// ---- 99_Test/PRG_TestPeakLive.TcPOU
PROGRAM PRG_TestPeakLive		// 피크컷(3)·통합(4) 모드 실제 경로 시험 (시험 모드, MAIN이 부름). bStart := TRUE로 시작, 약 10~15분
// 부하 모델: 가상 접속점 P = ESS 출력 − 부하 (수전 = 부하 − ESS 방전). 목표 피크 300 kW, 방전 허용 시간 끔 (PLC 시계 UTC)
// 피크컷: P1 부하 500 → 피크 방전, P2 부하 200 → 0, P3 자동 충전 시간 → 충전, P4 잔량 방전 시간 → 방전 (역송 방지 상한)
// 통합:   I1 부하 200·시간표 +100 → 100, I2 부하 600 → 피크·시간표 중 큰 값, I3 부하 200·시간표 −200 → 충전, I4 잔량 방전
// 구간마다 조건이 5 s 이어지면 통과·기록. 끝나면 설정·가상신호·운전 모드 되돌리고 PCS 정지
VAR
	bStart		: BOOL;				// TRUE로 쓰면 시작
	bDone		: BOOL;
	bPass		: BOOL;				// 8구간 모두 통과
	nStep		: UINT;
	wsStep		: WSTRING(80);		// 지금 단계
	wsFail		: WSTRING(80);
	(* 지금 값 *)
	fLoadSim	: REAL;				// kW, 모의 부하
	fImport		: REAL;				// kW, 수전 (= 부하 − ESS 출력)
	nActiveMode	: UINT;				// 3 = 피크컷, 4 = 통합
	nState		: UINT;				// 켜진 모드 상태 (GVL_CM_RSN: 0 정상, 11 피크, 12 피크 필요 없음, 13 자동 충전, 14 잔량 방전, 15 스케줄·피크, 6 역송 방지)
	fModeP		: REAL;				// 모드가 낸 값 (kW, 방전 +)
	fMgrP		: REAL;				// 관리자 지령
	fUnitP		: REAL;				// 가상 PCS 실제 출력
	fPeakCtrl	: REAL;				// 피크 제어량
	nRemainMin	: UINT;				// 15분 구간 남은 분
	fSoc		: REAL;				// %
	eRun		: E_RunState;
	stNow		: ST_LocalTime;
	(* 구간 결과 (통과 때 실제 출력 kW) *)
	bP1Peak		: BOOL;		fP1		: REAL;		// 피크컷: 부하 500 → 피크 방전
	bP2Below	: BOOL;		fP2		: REAL;		// 피크컷: 부하 200 → 0
	bP3AutoChg	: BOOL;		fP3		: REAL;		// 피크컷: 자동 충전
	bP4Remain	: BOOL;		fP4		: REAL;		// 피크컷: 잔량 방전
	bI1Sched	: BOOL;		fI1		: REAL;		// 통합: 시간표 +100
	bI2Peak		: BOOL;		fI2		: REAL;		// 통합: 피크·시간표 중 큰 값
	bI3Chg		: BOOL;		fI3		: REAL;		// 통합: 시간표 충전 −200
	bI4Remain	: BOOL;		fI4		: REAL;		// 통합: 잔량 방전
	(* 내부 *)
	bLoadSim	: BOOL;
	nLastStep	: UINT;
	tonStep		: TON;
	tonOk		: TON;
	bCond		: BOOL;
	bBackedUp	: BOOL;
	stCommonBak	: ST_CmCommonSet;
	stSchedBak	: ST_CmScheduleSet;
	stPeakBak	: ST_CmPeakCutSet;
	stSPBak		: ST_CmSchedPeakSet;
	stVirtBak	: ST_VirtualSet;
	stCmBak		: ST_CtrlModeSet;
	stMgrOut	: ST_SourceOutput;
	nMin		: UINT;
	nSeason		: UINT;
	k			: UINT;
	nWinStart	: UINT;		// HHMM
	nWinEnd		: UINT;		// HHMM (지금 + 3분)
	nSlotEnd	: UINT;		// HHMM (지금 + 30분)
END_VAR

// 지금 값
stNow		:= MAIN.fbClock.q_stTime;
nActiveMode	:= GVL_SITE.g_fbCtrlMode1.q_nActive;
stMgrOut	:= GVL_SITE.g_fbCtrlMode1.Output;
fMgrP		:= stMgrOut.fPSet;	// [16번 수정 2026-11-09: 관리자가 접속점 그룹 단위 → 접속점 그룹 지령 칸. 원래 stMgrOut.astUnit[1].fPSet (PCS2는 Manual이라 접속점 그룹 지령이 유닛 1로 감)]
fUnitP		:= MAIN.fbSnapshot.q_astUnit[1].stP.fValue;
eRun		:= MAIN.fbSnapshot.q_astUnit[1].eRunState;
fSoc		:= MAIN.fbGroupView.q_astView[1].stSocAvg.fValue;
IF nActiveMode = 4 THEN
	nState		:= GVL_SITE.g_fbCmSchedPeak1.q_nState;
	fModeP		:= GVL_SITE.g_fbCmSchedPeak1.q_fOutP;
	fPeakCtrl	:= GVL_SITE.g_fbCmSchedPeak1.q_fPeakCtrl;
	nRemainMin	:= GVL_SITE.g_fbCmSchedPeak1.q_nRemainMin;
ELSE
	nState		:= GVL_SITE.g_fbCmPeakCut1.q_nState;
	fModeP		:= GVL_SITE.g_fbCmPeakCut1.q_fOutP;
	fPeakCtrl	:= GVL_SITE.g_fbCmPeakCut1.q_fPeakCtrl;
	nRemainMin	:= GVL_SITE.g_fbCmPeakCut1.q_nRemainMin;
END_IF
// 부하 모델: 접속점 P (공급 +) = ESS 출력 − 부하
IF bLoadSim THEN
	GVL_TEST.g_astVirtual[1].bPEna	:= TRUE;
	GVL_TEST.g_astVirtual[1].fP		:= MAIN.fbGroupView.q_astView[1].fPOut - fLoadSim;	// 그룹 출력 (PCS2는 Manual 0)
END_IF
fImport := fLoadSim - fUnitP;
// 시간 구간 (지금 분 ~ +3분, 시간표 칸은 +30분)
nMin		:= stNow.nHour * 60 + stNow.nMinute;
nWinStart	:= (nMin / 60) * 100 + nMin MOD 60;
nWinEnd		:= (((nMin + 3) MOD 1440) / 60) * 100 + ((nMin + 3) MOD 1440) MOD 60;
nSlotEnd	:= (((nMin + 30) MOD 1440) / 60) * 100 + ((nMin + 30) MOD 1440) MOD 60;

tonStep(IN := nStep >= 20 AND nStep < 900, PT := T#240S);
bCond := FALSE;

CASE nStep OF
	0:
		IF bStart THEN
			bStart := FALSE;	bDone := FALSE;	bPass := FALSE;	wsFail := "";
			bP1Peak := FALSE;	bP2Below := FALSE;	bP3AutoChg := FALSE;	bP4Remain := FALSE;
			bI1Sched := FALSE;	bI2Peak := FALSE;	bI3Chg := FALSE;	bI4Remain := FALSE;
			nStep := 10;
		ELSIF NOT bDone THEN
			wsStep := "대기: bStart := TRUE로 시작";
		END_IF

	10:	// 준비
		wsStep := "설정 준비";
		IF NOT stNow.bValid OR stNow.nMonth < 1 OR stNow.nMonth > 12 OR stNow.nDay < 1 OR stNow.nDay > 31 OR stNow.nDayOfWeek > 6 THEN
			wsFail := "PLC 시각 무효";
			nStep := 900;
		ELSIF nMin + 40 >= 1440 THEN
			wsFail := "자정 가까움: 40분 뒤 다시";
			nStep := 900;
		ELSE
			stCommonBak	:= GVL_PERSIST.g_stModuleSet.stCmCommon;
			stSchedBak	:= GVL_PERSIST.g_stModuleSet.stCmSchedule1;
			stPeakBak	:= GVL_PERSIST.g_stModuleSet.stCmPeakCut1;
			stSPBak		:= GVL_PERSIST.g_stModuleSet.stCmSchedPeak1;
			stVirtBak	:= GVL_TEST.g_astVirtual[1];
			stCmBak		:= GVL_PERSIST.g_stModuleSet.stCtrlMode1;
			GVL_PERSIST.g_stModuleSet.stCtrlMode1.ePccShare := E_PccShare.Actual;	// PCS1이 접속점 실측 그대로 (PCS2는 Manual 0)
			bBackedUp	:= TRUE;
			GVL_PERSIST.g_stModuleSet.stCmCommon.stDis.bUse := FALSE;
			GVL_PERSIST.g_stModuleSet.stCmCommon.abHoliday[stNow.nMonth, stNow.nDay] := FALSE;
			GVL_PERSIST.g_stModuleSet.stCmPeakCut1.stPeak.fTarget	:= 300.0;
			GVL_PERSIST.g_stModuleSet.stCmPeakCut1.stAutoChg.bUse	:= FALSE;
			GVL_PERSIST.g_stModuleSet.stCmPeakCut1.stRemain.bUse		:= FALSE;
			GVL_PERSIST.g_stModuleSet.stCmSchedPeak1.stPeak.fTarget	:= 300.0;
			GVL_PERSIST.g_stModuleSet.stCmSchedPeak1.stRemain.bUse	:= FALSE;
			nSeason := GVL_PERSIST.g_stModuleSet.stCmCommon.anSeasonOfMonth[stNow.nMonth];
			IF nSeason > 2 THEN
				nSeason := 0;
			END_IF
			FOR k := 1 TO GVL_PARAM.SCHED_SLOT_COUNT DO
				GVL_PERSIST.g_stModuleSet.stCmSchedule1.astSlot[nSeason, stNow.nDayOfWeek, k].nStart	:= 0;
				GVL_PERSIST.g_stModuleSet.stCmSchedule1.astSlot[nSeason, stNow.nDayOfWeek, k].nEnd	:= 0;
				GVL_PERSIST.g_stModuleSet.stCmSchedule1.astSlot[nSeason, stNow.nDayOfWeek, k].fP		:= 0.0;
			END_FOR
			fLoadSim	:= 500.0;
			bLoadSim	:= TRUE;
			GVL_PERSIST.g_aeOpMode[1] := E_OpMode.Auto;
			nStep := 20;
		END_IF

	20:
		wsStep := "Auto 전환 대기";
		IF MAIN.fbModeSwitch.q_aeOpMode[1] = E_OpMode.Auto THEN
			GVL_SITE.g_fbSrcTest.i_nBatGroup	:= 0;
			GVL_SITE.g_fbSrcTest.i_eBatReq		:= E_BatCmd.Close;
			nStep := 30;
		END_IF
	30:
		wsStep := "배터리 투입 대기";
		IF MAIN.fbBatGroup.q_astBatGroup[1].bReady THEN
			GVL_SITE.g_fbSrcTest.i_nPcsUnit	:= 0;
			GVL_SITE.g_fbSrcTest.i_ePcsReq	:= E_PcsCmd.Run;
			nStep := 40;
		END_IF
	40:
		wsStep := "PCS Run 대기";
		IF eRun = E_RunState.Run THEN
			GVL_SITE.g_fbCtrlMode1.i_nModeReq := 3;
			nStep := 50;
		END_IF
	50:
		wsStep := "피크컷 모드 켜는 중";
		IF nActiveMode = 3 THEN
			nStep := 100;
		END_IF

	100: // P1 부하 500 > 목표 300 → 피크 방전
		wsStep := "P1 피크컷: 부하 500 > 목표 300";
		bCond := nActiveMode = 3 AND nState = GVL_CM_RSN.PEAK AND fPeakCtrl > 0.0 AND fModeP > 0.0 AND ABS(fUnitP - fModeP) < 5.0;
		IF tonOk.Q THEN
			bP1Peak := TRUE;	fP1 := fUnitP;
			fLoadSim := 200.0;
			nStep := 110;
		END_IF
	110: // P2 부하 200 < 목표 → 0
		wsStep := "P2 피크컷: 부하 200 < 목표 300";
		bCond := nState = GVL_CM_RSN.BELOW_PEAK AND ABS(fUnitP) < 5.0;
		IF tonOk.Q THEN
			bP2Below := TRUE;	fP2 := fUnitP;
			GVL_PERSIST.g_stModuleSet.stCmPeakCut1.stAutoChg.nStart	:= nWinStart;
			GVL_PERSIST.g_stModuleSet.stCmPeakCut1.stAutoChg.nEnd	:= nWinEnd;
			GVL_PERSIST.g_stModuleSet.stCmPeakCut1.stAutoChg.fSoc	:= 100.0;
			GVL_PERSIST.g_stModuleSet.stCmPeakCut1.stAutoChg.bUse	:= TRUE;
			nStep := 120;
		END_IF
	120: // P3 자동 충전 시간
		wsStep := "P3 피크컷: 자동 충전 시간";
		bCond := nState = GVL_CM_RSN.AUTO_CHG AND fModeP < -5.0 AND fUnitP < -5.0;
		IF tonOk.Q THEN
			bP3AutoChg := TRUE;	fP3 := fUnitP;
			GVL_PERSIST.g_stModuleSet.stCmPeakCut1.stAutoChg.bUse	:= FALSE;
			GVL_PERSIST.g_stModuleSet.stCmPeakCut1.stRemain.nStart	:= nWinStart;
			GVL_PERSIST.g_stModuleSet.stCmPeakCut1.stRemain.nEnd		:= nWinEnd;
			GVL_PERSIST.g_stModuleSet.stCmPeakCut1.stRemain.fSoc		:= 10.0;
			GVL_PERSIST.g_stModuleSet.stCmPeakCut1.stRemain.bUse		:= TRUE;
			fLoadSim := 500.0;
			nStep := 130;
		END_IF
	130: // P4 잔량 방전 시간 (역송 방지 상한)
		wsStep := "P4 피크컷: 잔량 방전 시간";
		bCond := (nState = GVL_CM_RSN.REMAIN_DIS OR nState = GVL_CM_RSN.REV_LIMIT) AND fModeP > 5.0 AND ABS(fUnitP - fModeP) < 5.0 AND fUnitP < fLoadSim;
		IF tonOk.Q THEN
			bP4Remain := TRUE;	fP4 := fUnitP;
			GVL_PERSIST.g_stModuleSet.stCmPeakCut1.stRemain.bUse := FALSE;
			// 통합 준비: 시간표 +100 (지금 ~ +30분), 부하 200
			GVL_PERSIST.g_stModuleSet.stCmSchedule1.astSlot[nSeason, stNow.nDayOfWeek, 1].nStart	:= nWinStart;
			GVL_PERSIST.g_stModuleSet.stCmSchedule1.astSlot[nSeason, stNow.nDayOfWeek, 1].nEnd	:= nSlotEnd;
			GVL_PERSIST.g_stModuleSet.stCmSchedule1.astSlot[nSeason, stNow.nDayOfWeek, 1].fP		:= 100.0;
			fLoadSim := 200.0;
			GVL_SITE.g_fbCtrlMode1.i_nModeReq := 4;
			nStep := 200;
		END_IF

	200:
		wsStep := "통합 모드 켜는 중";
		IF nActiveMode = 4 THEN
			nStep := 210;
		END_IF
	210: // I1 부하 200 (피크 아님) → 시간표 +100
		wsStep := "I1 통합: 부하 200, 시간표 +100";
		bCond := nState = 0 AND ABS(fModeP - 100.0) < 0.5 AND ABS(fUnitP - 100.0) < 5.0;
		IF tonOk.Q THEN
			bI1Sched := TRUE;	fI1 := fUnitP;
			fLoadSim := 600.0;
			nStep := 220;
		END_IF
	220: // I2 부하 600 > 목표 → 피크 제어량과 시간표 중 큰 값
		wsStep := "I2 통합: 부하 600 > 목표 300";
		bCond := nState = GVL_CM_RSN.SCHED_PEAK AND fPeakCtrl > 0.0 AND fModeP >= 99.9 AND ABS(fModeP - MAX(fPeakCtrl, 100.0)) < 0.5 AND ABS(fUnitP - fModeP) < 5.0;
		IF tonOk.Q THEN
			bI2Peak := TRUE;	fI2 := fUnitP;
			GVL_PERSIST.g_stModuleSet.stCmSchedule1.astSlot[nSeason, stNow.nDayOfWeek, 1].fP := -200.0;
			fLoadSim := 200.0;
			nStep := 230;
		END_IF
	230: // I3 부하 200, 시간표 충전 −200
		wsStep := "I3 통합: 부하 200, 시간표 -200";
		bCond := nState = 0 AND ABS(fModeP + 200.0) < 0.5 AND ABS(fUnitP + 200.0) < 5.0;
		IF tonOk.Q THEN
			bI3Chg := TRUE;	fI3 := fUnitP;
			GVL_PERSIST.g_stModuleSet.stCmSchedPeak1.stRemain.nStart	:= nWinStart;
			GVL_PERSIST.g_stModuleSet.stCmSchedPeak1.stRemain.nEnd	:= nWinEnd;
			GVL_PERSIST.g_stModuleSet.stCmSchedPeak1.stRemain.fSoc	:= 10.0;
			GVL_PERSIST.g_stModuleSet.stCmSchedPeak1.stRemain.bUse	:= TRUE;
			fLoadSim := 500.0;
			nStep := 240;
		END_IF
	240: // I4 잔량 방전
		wsStep := "I4 통합: 잔량 방전 시간";
		bCond := (nState = GVL_CM_RSN.REMAIN_DIS OR nState = GVL_CM_RSN.REV_LIMIT) AND fModeP > 5.0 AND ABS(fUnitP - fModeP) < 5.0 AND fUnitP < fLoadSim;
		IF tonOk.Q THEN
			bI4Remain := TRUE;	fI4 := fUnitP;
			nStep := 900;
		END_IF

	900: // 정리
		GVL_SITE.g_fbCtrlMode1.i_nModeReq	:= 0;
		GVL_SITE.g_fbSrcTest.i_nPcsUnit		:= 0;
		GVL_SITE.g_fbSrcTest.i_ePcsReq		:= E_PcsCmd.Stop;
		bLoadSim := FALSE;
		IF bBackedUp THEN
			GVL_PERSIST.g_stModuleSet.stCmCommon	:= stCommonBak;
			GVL_PERSIST.g_stModuleSet.stCmSchedule1	:= stSchedBak;
			GVL_PERSIST.g_stModuleSet.stCmPeakCut1	:= stPeakBak;
			GVL_PERSIST.g_stModuleSet.stCmSchedPeak1	:= stSPBak;
			GVL_TEST.g_astVirtual[1]				:= stVirtBak;
			GVL_PERSIST.g_stModuleSet.stCtrlMode1	:= stCmBak;
			bBackedUp := FALSE;
		END_IF
		GVL_PERSIST.g_aeOpMode[1] := E_OpMode.Manual;
		bPass := bP1Peak AND bP2Below AND bP3AutoChg AND bP4Remain AND bI1Sched AND bI2Peak AND bI3Chg AND bI4Remain AND wsFail = "";
		bDone := TRUE;
		IF bPass THEN
			wsStep := "끝: 통과";
		ELSE
			wsStep := "끝: 실패 (wsFail·구간 결과 확인)";
		END_IF
		nStep := 0;
END_CASE

// 조건이 5 s 이어지면 통과 (단계가 바뀌면 다시 셈)
tonOk(IN := bCond AND nStep = nLastStep, PT := T#5S);
IF tonStep.Q AND nStep >= 20 AND nStep < 900 THEN
	wsFail	:= WCONCAT("시간 초과: ", wsStep);
	nStep	:= 900;
END_IF
IF nStep <> nLastStep THEN
	tonStep(IN := FALSE);
	tonOk(IN := FALSE);
	nLastStep := nStep;
END_IF

END_PROGRAM

// ---- 99_Test/PRG_TestUnitMode.TcPOU
PROGRAM PRG_TestUnitMode		// PCS별(유닛 단위) 제어 모드 자동 시험 (GVL_SITE.TEST_MODE일 때 MAIN이 부름). 따로 둔 인스턴스만 씀 (장비 지령에 영향 없음)
// 온라인에서 bDone = TRUE가 되면 fbTally.q_nPass·q_nFail, 실패하면 fbTally.q_anFail. bRestart := TRUE로 다시 돌림
// 40~41: 유닛 단위 출력 칸, 42~44: 접속점 몫 (ByRating·Actual·Fixed), 45~47: 설정 점검, 48~50: FB_UnitView 버스 몫, 51~57: 스탠다드 스케줄 모드, 58~63: NaN·무한대 거르기 (PLC가 멈추지 않아야 함)
VAR
	bRestart	: BOOL;
	bDone		: BOOL;
	nStep		: UINT;
	fbTally		: FB_TestTally;
	fbConstU	: FB_CmConstPower	:= (i_nModuleId := 9012, i_sName := 'TestConstU');
	fbMgrU		: FB_CtrlModeMgr	:= (i_nModuleId := 9010, i_sName := 'TestMgrU', i_nUnit := 1);
	aipMode		: ARRAY[1..GVL_PARAM.CTRL_MODE_COUNT] OF I_ControlMode;
	astUv		: ARRAY[1..GVL_PARAM.UNIT_COUNT] OF ST_UnitView;	// 관리자에 주소로 넘기는 유닛 값 (시험이 채움)
	stGrpView	: ST_GroupView;			// 지령원 공통 입력 (유닛 단위에서는 안 봄)
	stReg		: ST_SourceReg := (bEnable := TRUE, nGrade := 1, ePowerMode := E_SourceMode.Auto, nGroup := 0, tExpire := T#10S);
	stMgrOut	: ST_SourceOutput;
	wsTmp		: WSTRING(63);
	(* FB_UnitView 시험 (유닛 1 기준, 유닛이 2개 이상이면 유닛 2도) *)
	fbUv		: FB_UnitView;
	astView		: ARRAY[1..GVL_PARAM.GROUP_COUNT] OF ST_GroupView;
	astUnit		: ARRAY[1..GVL_PARAM.UNIT_COUNT] OF ST_UnitState;
	astAvail	: ARRAY[1..GVL_PARAM.UNIT_COUNT] OF ST_UnitAvail;
	astCfg		: ARRAY[1..GVL_PARAM.UNIT_COUNT] OF ST_UnitCfg;
	astEnv		: ARRAY[1..GVL_PARAM.UNIT_COUNT] OF ST_UnitEnvelope;
	astBat		: ARRAY[1..GVL_PARAM.BAT_COUNT] OF ST_BatGroupState;
	astBatEnv	: ARRAY[1..GVL_PARAM.BAT_COUNT] OF ST_BatEnvelope;
	fShareExp	: REAL;
	(* 스탠다드 스케줄 모드 시험 *)
	fbStd		: FB_CmStdSchedule	:= (i_nModuleId := 9013, i_sName := 'TestStdSched');
	stStdView	: ST_CtrlModeView;
	stStdOut	: ST_CtrlModeOut;
	nInfBits	: DWORD := 16#7F800000;	// +무한대 비트 (NaN은 크기 비교에서 부동소수점 예외로 PLC가 멈추므로 시험에 쓰지 않음)
	fInf		: REAL;
	nBad0		: UDINT;
	nNanBits	: DWORD := 16#7FC00000;	// NaN 비트 (거르기 시험: 비교하기 전에 걸러져야 PLC가 멈추지 않음)
	fNan		: REAL;
	fbEmsCmd	: FB_EmsCommand;		// EMS 명령 핸들러 시험 인스턴스
	astPcsRx	: ARRAY[0..GVL_PARAM.PCS_COUNT - 1] OF ST_MqttCommand_Rx;
	astBatRx	: ARRAY[0..GVL_PARAM.BMS_COUNT - 1] OF ST_MqttCommand_Rx;
	nPSeq0		: UDINT;
	nRunSeq0	: UDINT;		// 시험 전 이상값 버린 수 (누계라 다시 돌려도 맞게)
	u			: UINT;
END_VAR

IF bRestart THEN
	bRestart	:= FALSE;
	bDone		:= FALSE;
	nStep		:= 0;
END_IF

CASE nStep OF
	0:	// 준비: 정출력 80 kW 하나, 유닛 1 값 (출력 100, 그룹 출력 300, 접속점 -200 = 수전 200 → 그룹 부하 500, 몫 0.5)
		fbTally.M_Reset();
		aipMode[1]					:= fbConstU;
		fbConstU.i_stSet.fPSet		:= 80.0;
		fbConstU.i_stSet.bQSet		:= FALSE;
		fbConstU.i_stSet.tDuration	:= T#0S;
		astUv[1].nUnit				:= 1;
		astUv[1].bAvail				:= TRUE;
		astUv[1].stView.nUnitAvail	:= 1;
		astUv[1].stView.fPRatedAvail	:= 1000.0;
		astUv[1].stView.fPOut		:= 100.0;
		astUv[1].stView.stPcc.stMeas.stP.bValid	:= TRUE;
		astUv[1].stView.stPcc.stMeas.stP.fValue	:= -200.0;
		astUv[1].fGroupPOut			:= 300.0;
		astUv[1].fRatingShare		:= 0.5;
		fbMgrU.i_aipMode			:= aipMode;
		fbMgrU.i_stSet.bZeroOnSwitch	:= TRUE;
		fbMgrU.i_stSet.tZeroDelay	:= T#1S;
		fbMgrU.i_stSet.nFallback	:= 0;
		fbMgrU.i_stSet.ePccShare	:= E_PccShare.ByRating;
		fbMgrU.i_stSet.fPccRatio	:= 1.0;
		fbMgrU.i_pUnitView			:= ADR(astUv);
		wsTmp := fbMgrU.M_CheckSet();
		fbTally.M_Check(i_nId := 40, i_bOk := wsTmp = "");
		fbMgrU.i_nModeReq := 1;
		nStep := 10;

	10:	// 정출력 진입: 유닛 1 칸에만 80, 그룹 지령은 없음. 몫 0.5 → 모드가 본 접속점 = 100 - 0.5 × 500 = -150
		A_Cycle();
		fbTally.M_Check(i_nId := 41, i_bOk := fbMgrU.q_nActive = 1 AND stMgrOut.astUnit[1].bPSetActive AND ABS(stMgrOut.astUnit[1].fPSet - 80.0) < 0.01 AND NOT stMgrOut.bPSetActive);
		fbTally.M_Check(i_nId := 42, i_bOk := ABS(fbMgrU.q_fPccP + 150.0) < 0.01);
		fbMgrU.i_stSet.ePccShare := E_PccShare.Actual;
		nStep := 11;

	11:	// Actual: 실측 그대로 -200
		A_Cycle();
		fbTally.M_Check(i_nId := 43, i_bOk := ABS(fbMgrU.q_fPccP + 200.0) < 0.01);
		fbMgrU.i_stSet.ePccShare := E_PccShare.Fixed;
		fbMgrU.i_stSet.fPccRatio := 0.2;
		nStep := 12;

	12:	// Fixed 0.2: 100 - 0.2 × 500 = 0
		A_Cycle();
		fbTally.M_Check(i_nId := 44, i_bOk := ABS(fbMgrU.q_fPccP) < 0.01);
		// 설정 점검: 몫 범위 밖, 유닛 값 연결 안 됨, 유닛 번호 범위 밖
		fbMgrU.i_stSet.fPccRatio := 1.5;
		wsTmp := fbMgrU.M_CheckSet();
		fbTally.M_Check(i_nId := 45, i_bOk := wsTmp <> "");
		fbMgrU.i_stSet.fPccRatio := 0.2;
		fbMgrU.i_pUnitView := 0;
		wsTmp := fbMgrU.M_CheckSet();
		fbTally.M_Check(i_nId := 46, i_bOk := wsTmp <> "");
		fbMgrU.i_pUnitView := ADR(astUv);
		fbMgrU.i_nUnit := GVL_PARAM.UNIT_COUNT + 1;
		wsTmp := fbMgrU.M_CheckSet();
		fbTally.M_Check(i_nId := 47, i_bOk := wsTmp <> "");
		fbMgrU.i_nUnit := 1;
		A_UnitViewTest();
		A_StdScheduleTest();
		A_NanTest();
		nStep := 99;

	99:
		bDone := TRUE;
END_CASE

ACTION A_Cycle:
fbMgrU.i_pUnitView := ADR(astUv);	// 온라인 변경 뒤에도 맞게 매번
fbMgrU.M_Cycle(i_stReg := stReg, i_stView := stGrpView);
stMgrOut := fbMgrU.Output;
END_ACTION

ACTION A_UnitViewTest:
// FB_UnitView: 그룹 1 (접속점 -200, 그룹 출력 300, 가용 한도 합 2000), 버스 1 (방전 한도 1200, 충전 한도 800, 용량 4000, SOC 60)
// 유닛 1 정격 1000 (한도 1000, 출력 100). 유닛이 2개 이상이면 유닛 2도 같은 버스·정격 1000 → 버스 몫 0.5, 아니면 1
astView[1].stPcc.stMeas.stP.bValid	:= TRUE;
astView[1].stPcc.stMeas.stP.fValue	:= -200.0;
astView[1].fPOut			:= 300.0;
astView[1].fPRatedAvail		:= 2000.0;
astBat[1].bUsable			:= TRUE;
astBat[1].fCapacity			:= 4000.0;
astBat[1].stSoc.bValid		:= TRUE;
astBat[1].stSoc.fValue		:= 60.0;
astBatEnv[1].stP.fMax		:= 1200.0;
astBatEnv[1].stP.fMin		:= -800.0;
FOR u := 1 TO GVL_PARAM.UNIT_COUNT DO
	astCfg[u].nGroup		:= 1;
	astCfg[u].nBatGroup		:= 1;
	astCfg[u].fPRated		:= 1000.0;
	astCfg[u].fQRated		:= 500.0;
	astAvail[u].bAvail		:= TRUE;
	astEnv[u].stP.fMax		:= 1000.0;
	astEnv[u].stQ.fMax		:= 500.0;
	astUnit[u].stP.bValid	:= TRUE;
	astUnit[u].stP.fValue	:= 100.0;
END_FOR
fShareExp := 1.0 / UINT_TO_REAL(GVL_PARAM.UNIT_COUNT);
fbUv(iq_astView := astView, iq_astUnit := astUnit, iq_astAvail := astAvail, iq_astUnitCfg := astCfg,
	iq_astUnitEnv := astEnv, iq_astBatGroup := astBat, iq_astBatEnv := astBatEnv);
// 48) 유닛 1: 출력·한도·접속점·그룹 출력·정격 몫 (1000 / 2000)
fbTally.M_Check(i_nId := 48, i_bOk := fbUv.q_astView[1].stView.nUnitAvail = 1 AND ABS(fbUv.q_astView[1].stView.fPOut - 100.0) < 0.01
	AND ABS(fbUv.q_astView[1].stView.fPRatedAvail - 1000.0) < 0.01 AND ABS(fbUv.q_astView[1].stView.stPcc.stMeas.stP.fValue + 200.0) < 0.01
	AND ABS(fbUv.q_astView[1].fGroupPOut - 300.0) < 0.01 AND ABS(fbUv.q_astView[1].fRatingShare - 0.5) < 0.001);
// 49) 버스 몫: 용량·방전·충전 한도 × 몫, SOC 그대로
fbTally.M_Check(i_nId := 49, i_bOk := ABS(fbUv.q_astView[1].stView.fCapacity - 4000.0 * fShareExp) < 0.1
	AND ABS(fbUv.q_astView[1].stView.fPDisMax - MIN(1200.0 * fShareExp, 1000.0)) < 0.1 AND ABS(fbUv.q_astView[1].stView.fPChgMax - MIN(800.0 * fShareExp, 1000.0)) < 0.1
	AND fbUv.q_astView[1].stView.stSocAvg.bValid AND ABS(fbUv.q_astView[1].stView.stSocAvg.fValue - 60.0) < 0.01);
// 50) 가용이 아닌 유닛: 가용 0, 몫 0, 용량 0
astAvail[1].bAvail := FALSE;
fbUv(iq_astView := astView, iq_astUnit := astUnit, iq_astAvail := astAvail, iq_astUnitCfg := astCfg,
	iq_astUnitEnv := astEnv, iq_astBatGroup := astBat, iq_astBatEnv := astBatEnv);
fbTally.M_Check(i_nId := 50, i_bOk := fbUv.q_astView[1].stView.nUnitAvail = 0 AND fbUv.q_astView[1].fRatingShare = 0.0 AND fbUv.q_astView[1].stView.fCapacity = 0.0
	AND ABS(fbUv.q_astView[1].stView.fPOut - 100.0) < 0.01);
astAvail[1].bAvail := TRUE;
END_ACTION

ACTION A_StdScheduleTest:
// 스탠다드 스케줄: EMS가 9시 방전 100, 10시 정지를 보내는 흐름 (한 스캔씩 직접 부름)
stStdView.stGroup.nUnitAvail := 1;
// 켜지기 전에 온 지령(번호 5, 50 kW)은 쓰지 않음
fbStd.i_astCmd[1].bUse		:= TRUE;	// [16번 수정 2026-11-09: 모드가 유닛마다 칸을 받음 (유닛 1 칸으로 시험). 원래 fbStd.i_stCmd, 출력 stStdOut.bPSetActive·fPSet]
fbStd.i_astCmd[1].bAlive	:= TRUE;
fbStd.i_astCmd[1].nPSeq		:= 5;
fbStd.i_astCmd[1].fP		:= 50.0;
fbStd.i_astCmd[1].nStateSeq	:= 3;
fbStd.i_astCmd[1].eState	:= E_PcsCmd.Run;
fbStd.M_Enter(i_stView := stStdView);
stStdOut := fbStd.M_Calc(i_stView := stStdView);
fbTally.M_Check(i_nId := 51, i_bOk := stStdOut.bUnitOut AND stStdOut.astUnit[1].bPSetActive AND stStdOut.astUnit[1].fPSet = 0.0 AND fbStd.q_nState = 3 AND NOT fbStd.q_abHold[1]);
// 9시: 방전 100 → 100, 다음 지령까지 유지
fbStd.i_astCmd[1].nPSeq	:= 6;
fbStd.i_astCmd[1].fP	:= 100.0;
stStdOut := fbStd.M_Calc(i_stView := stStdView);
stStdOut := fbStd.M_Calc(i_stView := stStdView);
fbTally.M_Check(i_nId := 52, i_bOk := ABS(stStdOut.astUnit[1].fPSet - 100.0) < 0.01 AND fbStd.q_nState = 0 AND fbStd.q_nCmdCount = 1);
// 10시: 정지 → 0 (새 P 지령 대기)
fbStd.i_astCmd[1].nStateSeq	:= 4;
fbStd.i_astCmd[1].eState	:= E_PcsCmd.Stop;
stStdOut := fbStd.M_Calc(i_stView := stStdView);
fbTally.M_Check(i_nId := 53, i_bOk := stStdOut.astUnit[1].bPSetActive AND stStdOut.astUnit[1].fPSet = 0.0 AND fbStd.q_nState = 3);
// Run만 다시 와도 옛 100은 되살아나지 않음
fbStd.i_astCmd[1].nStateSeq	:= 5;
fbStd.i_astCmd[1].eState	:= E_PcsCmd.Run;
stStdOut := fbStd.M_Calc(i_stView := stStdView);
fbTally.M_Check(i_nId := 54, i_bOk := stStdOut.astUnit[1].fPSet = 0.0 AND NOT fbStd.q_abHold[1]);
// 충전 -200 → -200. 이상값(무한대)은 버리고 앞 값 유지
fbStd.i_astCmd[1].nPSeq	:= 7;
fbStd.i_astCmd[1].fP	:= -200.0;
stStdOut := fbStd.M_Calc(i_stView := stStdView);
nBad0 := fbStd.q_nBadCount;
fbStd.i_astCmd[1].nPSeq	:= 8;
MEMCPY(destAddr := ADR(fInf), srcAddr := ADR(nInfBits), n := SIZEOF(fInf));	// +무한대 (비트로 만듦)
fbStd.i_astCmd[1].fP	:= fInf;
stStdOut := fbStd.M_Calc(i_stView := stStdView);
fbTally.M_Check(i_nId := 55, i_bOk := ABS(stStdOut.astUnit[1].fPSet + 200.0) < 0.01 AND fbStd.q_nBadCount = nBad0 + 1);
// EMS 끊김 → 0, 돌아와도 옛 값은 되살아나지 않음
fbStd.i_astCmd[1].bAlive := FALSE;
stStdOut := fbStd.M_Calc(i_stView := stStdView);
fbTally.M_Check(i_nId := 56, i_bOk := stStdOut.astUnit[1].fPSet = 0.0 AND fbStd.q_nState = 2);
fbStd.i_astCmd[1].bAlive := TRUE;
stStdOut := fbStd.M_Calc(i_stView := stStdView);
fbTally.M_Check(i_nId := 57, i_bOk := stStdOut.astUnit[1].fPSet = 0.0 AND fbStd.q_nState = 3);
fbStd.M_Exit();
END_ACTION

ACTION A_NanTest:
// NaN·무한대: 비트로 먼저 거르는지 (거르지 못하면 여기서 PLC가 멈춤)
MEMCPY(destAddr := ADR(fNan), srcAddr := ADR(nNanBits), n := SIZEOF(fNan));
// 58) F_IsFinite: NaN·무한대 FALSE, 보통 숫자 TRUE
fbTally.M_Check(i_nId := 58, i_bOk := NOT F_IsFinite(fNan) AND NOT F_IsFinite(fInf) AND F_IsFinite(-123.4) AND F_IsFinite(0.0));
// 59) F_CmdOk: NaN은 한도가 있든 없든 FALSE, 보통 숫자는 한도대로
fbTally.M_Check(i_nId := 59, i_bOk := NOT F_CmdOk(fNan, 0.0) AND NOT F_CmdOk(fNan, 1000.0) AND NOT F_CmdOk(fInf, 0.0)
	AND F_CmdOk(500.0, 1000.0) AND NOT F_CmdOk(1500.0, 1000.0));
// 60) 스탠다드 스케줄 모드: NaN P 지령은 버리고 앞 값 유지
fbStd.i_astCmd[1].bAlive	:= TRUE;
fbStd.M_Enter(i_stView := stStdView);
fbStd.i_astCmd[1].nPSeq		:= fbStd.i_astCmd[1].nPSeq + 1;
fbStd.i_astCmd[1].fP		:= 70.0;
stStdOut := fbStd.M_Calc(i_stView := stStdView);
nBad0 := fbStd.q_nBadCount;
fbStd.i_astCmd[1].nPSeq		:= fbStd.i_astCmd[1].nPSeq + 1;
fbStd.i_astCmd[1].fP		:= fNan;
stStdOut := fbStd.M_Calc(i_stView := stStdView);
fbTally.M_Check(i_nId := 60, i_bOk := ABS(stStdOut.astUnit[1].fPSet - 70.0) < 0.01 AND fbStd.q_nBadCount = nBad0 + 1);
fbStd.M_Exit();
// 61) EMS 명령 핸들러: 방전 NaN → 버리고 셈, P 번호 안 바뀜 (PCS1 = 칸 0)
nPSeq0 := fbEmsCmd.q_stCmd.anPcsPSeq[1];
nBad0 := fbEmsCmd.q_nBadValueCount;
astPcsRx[0].Value		:= fNan;
astPcsRx[0].CommandType	:= 5;
fbEmsCmd(i_nRxCount := 1, iq_astPcsCommand := astPcsRx, iq_astBatCommand := astBatRx);
fbTally.M_Check(i_nId := 61, i_bOk := fbEmsCmd.q_nBadValueCount = nBad0 + 1 AND fbEmsCmd.q_stCmd.anPcsPSeq[1] = nPSeq0 AND astPcsRx[0].CommandType = 0);
// 62) 상태 명령(Run)에 Value가 NaN이어도 명령은 받음 (값은 안 봄)
nRunSeq0 := fbEmsCmd.q_stCmd.astPcs[1].nSeq;
astPcsRx[0].Value		:= fNan;
astPcsRx[0].CommandType	:= 1;
fbEmsCmd(i_nRxCount := 2, iq_astPcsCommand := astPcsRx, iq_astBatCommand := astBatRx);
fbTally.M_Check(i_nId := 62, i_bOk := fbEmsCmd.q_stCmd.astPcs[1].nSeq = nRunSeq0 + 1 AND fbEmsCmd.q_stCmd.astPcs[1].eCmd = E_PcsCmd.Run);
// 63) 보통 값(방전 120)은 받음
astPcsRx[0].Value		:= 120.0;
astPcsRx[0].CommandType	:= 5;
fbEmsCmd(i_nRxCount := 3, iq_astPcsCommand := astPcsRx, iq_astBatCommand := astBatRx);
fbTally.M_Check(i_nId := 63, i_bOk := fbEmsCmd.q_stCmd.anPcsPSeq[1] = nPSeq0 + 1 AND ABS(fbEmsCmd.q_stCmd.afPcsP[1] - 120.0) < 0.01);
END_ACTION

END_PROGRAM

// ---- 20_Module/ControlMode/FB_CmStdSchedule.TcPOU
FUNCTION_BLOCK FB_CmStdSchedule EXTENDS FB_CtrlModeBase		// 제어 모드: 스탠다드 스케줄. 시간표를 PMS에 두지 않고 EMS가 시각마다 보내는 지령을 그대로 따름
// 예) 09~10시 방전 100 kW: EMS가 9시에 방전 100 kW, 10시에 정지를 보냄 → 이 모드는 받은 P를 다음 지령까지 유지하고, 정지 쪽 명령이 오면 버림
// Manual 지령과 같은 구조: 새 지령(번호가 바뀜)만 받음, 받은 값은 다음 지령까지 유지, 정지 쪽 명령 뒤에는 새 P 지령이 올 때까지 0
//   - 모드가 켜지기 전에 온 지령은 쓰지 않음 (켜진 뒤 새 지령부터). 켜져 있는 동안 P는 늘 냄 (지령이 없으면 0 → 등급이 낮은 다른 지령원 값이 새지 않게)
//   - EMS가 끊기면 받아 둔 P를 버리고 0. 이상값(NaN·무한대)은 버리고 앞 값을 유지 (정격 대비 상한은 코어 명령 필터)
//   - 상태 명령(Run·Stop 등) 자체는 EMS 지령원(FB_SrcEms)이 장비에 냄. 이 모드는 P만 냄. 역송 방지·방전 허용 시간은 걸지 않음 (EMS 책임, 코어 접속점 제한은 그대로)
// [16번 수정 2026-11-09: 유닛마다 따로 받고 유닛별 값(bUnitOut)으로 냄. 제어 모드 관리자가 접속점 그룹 단위여도 EMS가 PCS마다 보낸 값을 그대로 따름.
//   원래는 PCS마다 관리자·모드 인스턴스(g_fbCmStdSched1·2)가 있고 지령 하나(i_stCmd)를 그 관리자 단위 값으로 냄]
// 입력 i_astCmd는 MAIN(A_PassEmsCmd)이 매 스캔 채움 (PCS 지령을 그 PCS의 유닛에 정격 비율로 나눔)
VAR_INPUT
	i_astCmd	: ARRAY[1..GVL_PARAM.UNIT_COUNT] OF ST_CmExtCmd;	// 유닛마다 바깥 지령. bUse FALSE인 칸은 내지 않음
END_VAR
VAR_OUTPUT
	q_nState	: UINT;				// 요약: 0 = 쓰는 유닛 모두 받은 P를 냄, 그 외 = 0을 내는 유닛의 첫 이유 (M_ReasonText)
	q_anState	: ARRAY[1..GVL_PARAM.UNIT_COUNT] OF UINT;	// 유닛마다 0 = 받은 P를 냄, 그 외 = 0을 내는 이유
	q_abHold	: ARRAY[1..GVL_PARAM.UNIT_COUNT] OF BOOL;	// 받아 둔 P 지령 있음
	q_afPCmd	: ARRAY[1..GVL_PARAM.UNIT_COUNT] OF REAL;	// kW, 받아 둔 P 지령 (q_abHold일 때)
	q_nCmdCount	: UDINT;			// 켜진 뒤 받은 P 지령 수 (유닛 합)
	q_nBadCount	: UDINT;			// 이상값이라 버린 P 지령 수
END_VAR
VAR
	_anPSeq		: ARRAY[1..GVL_PARAM.UNIT_COUNT] OF UDINT;	// 처리한 P 지령 번호
	_anStateSeq	: ARRAY[1..GVL_PARAM.UNIT_COUNT] OF UDINT;	// 처리한 상태 명령 번호
END_VAR
VAR CONSTANT
	RSN_NO_UNIT		: UINT := 1;	// 진입 거부: 가용 유닛 없음
	RSN_NO_EXT		: UINT := 2;	// EMS 끊김 → 0
	RSN_WAIT_CMD	: UINT := 3;	// 새 P 지령 대기 (켜진 뒤 아직 없음, 또는 정지 쪽 명령 뒤) → 0
END_VAR

METHOD M_CheckEnter : UINT
VAR_INPUT
	i_stView	: ST_CtrlModeView;	// 그룹 값(stGroup)·현지 시각(stTime). 관리자가 매 스캔 채움
END_VAR
M_CheckEnter := 0;
IF i_stView.stGroup.nUnitAvail = 0 THEN
	M_CheckEnter := RSN_NO_UNIT;
END_IF
END_METHOD

METHOD M_Enter
VAR_INPUT
	i_stView	: ST_CtrlModeView;	// 그룹 값(stGroup)·현지 시각(stTime). 관리자가 매 스캔 채움
END_VAR
VAR
	u			: UINT;
END_VAR
SUPER^.M_Enter(i_stView := i_stView);
// 켜지기 전에 온 지령은 쓰지 않음: 지금 번호를 처리한 것으로 두고 새 지령을 기다림
FOR u := 1 TO GVL_PARAM.UNIT_COUNT DO
	_anPSeq[u]		:= i_astCmd[u].nPSeq;
	_anStateSeq[u]	:= i_astCmd[u].nStateSeq;
	q_abHold[u]		:= FALSE;
	q_afPCmd[u]		:= 0.0;
END_FOR
q_nCmdCount	:= 0;
END_METHOD

METHOD M_Calc : ST_CtrlModeOut
VAR_INPUT
	i_stView	: ST_CtrlModeView;	// 그룹 값(stGroup)·현지 시각(stTime). 관리자가 매 스캔 채움
END_VAR
VAR
	u			: UINT;
	bNewCmd		: BOOL;		// 이번 스캔에 새 지령이 옴 (살아 있다는 표시)
	bAlive		: BOOL;
END_VAR
q_nState := 0;
FOR u := 1 TO GVL_PARAM.UNIT_COUNT DO
	bNewCmd := i_astCmd[u].nStateSeq <> _anStateSeq[u] OR i_astCmd[u].nPSeq <> _anPSeq[u];
	// 1) 상태 명령: 정지 쪽이면 받아 둔 P를 버림 (같은 메시지에 P가 같이 오면 아래에서 P가 다시 들어감)
	IF i_astCmd[u].nStateSeq <> _anStateSeq[u] THEN
		_anStateSeq[u] := i_astCmd[u].nStateSeq;
		IF i_astCmd[u].eState = E_PcsCmd.Stop OR i_astCmd[u].eState = E_PcsCmd.Standby OR i_astCmd[u].eState = E_PcsCmd.EStop THEN
			q_abHold[u] := FALSE;
		END_IF
	END_IF
	// 2) 새 P 지령: 다음 지령까지 유지. 이상값은 버리고 앞 값 유지
	IF i_astCmd[u].nPSeq <> _anPSeq[u] THEN
		_anPSeq[u] := i_astCmd[u].nPSeq;
		IF F_CmdOk(i_fValue := i_astCmd[u].fP, i_fLimit := 0.0) THEN
			q_abHold[u]	:= TRUE;
			q_afPCmd[u]	:= i_astCmd[u].fP;
			q_nCmdCount	:= q_nCmdCount + 1;
		ELSE
			q_nBadCount	:= q_nBadCount + 1;
		END_IF
	END_IF
	// 3) EMS가 끊기면 버림 (돌아와도 옛 지령이 되살아나지 않음).
	//    bAlive는 지난 스캔 값이라, 조용하던 EMS의 첫 지령 스캔에는 아직 FALSE → 새 지령이 온 스캔은 살아 있는 것으로 봄
	bAlive := i_astCmd[u].bAlive OR bNewCmd;
	IF NOT bAlive THEN
		q_abHold[u] := FALSE;
	END_IF
	// 4) 유닛 상태·출력: 쓰는 유닛은 켜져 있는 동안 P를 늘 냄. Q는 다른 지령원에 맡김
	IF q_abHold[u] THEN
		q_anState[u] := 0;
	ELSIF NOT bAlive THEN
		q_anState[u] := RSN_NO_EXT;
	ELSE
		q_anState[u] := RSN_WAIT_CMD;
	END_IF
	M_Calc.astUnit[u].bPSetActive	:= i_astCmd[u].bUse;
	M_Calc.astUnit[u].fPSet			:= SEL(q_abHold[u], 0.0, q_afPCmd[u]);
	M_Calc.astUnit[u].bQSetActive	:= FALSE;
	M_Calc.astUnit[u].fQSet			:= 0.0;
	IF i_astCmd[u].bUse AND q_nState = 0 THEN
		q_nState := q_anState[u];
	END_IF
END_FOR
M_Calc.bUnitOut		:= TRUE;		// 접속점 그룹 값(bPSetActive·fPSet)은 쓰지 않음
M_Calc.bPSetActive	:= FALSE;
M_Calc.fPSet		:= 0.0;
M_Calc.bQSetActive	:= FALSE;
M_Calc.fQSet		:= 0.0;
M_Calc.bExitReq		:= FALSE;
M_Calc.nReason		:= q_nState;
END_METHOD

METHOD M_ReasonText : WSTRING(63)
VAR_INPUT
	i_nReason	: UINT;
END_VAR
CASE i_nReason OF
	RSN_NO_UNIT:	M_ReasonText := "스탠다드 스케줄: 가용 유닛 없음";
	RSN_NO_EXT:		M_ReasonText := "스탠다드 스케줄: EMS 끊김 (0)";
	RSN_WAIT_CMD:	M_ReasonText := "스탠다드 스케줄: 새 P 지령 대기 (0)";
ELSE
	M_ReasonText := WCONCAT("이유 ", TO_WSTRING(i_nReason));
END_CASE
END_METHOD

END_FUNCTION_BLOCK

// ---- 99_Test/PRG_TestStdLive.TcPOU
PROGRAM PRG_TestStdLive		// 스탠다드 스케줄 모드 실제 경로 시험 (시험 모드, MAIN이 부름): EMS 명령 레코드 → FB_EmsCommand(MqttTask) → GVL_IF → MAIN A_PassEmsCmd → 모드 → 관리자 → 코어 고르기
// bStart := TRUE로 시작. PCS2(유닛 2)를 Auto로 두고 접속점 그룹 관리자(g_fbCtrlMode1)에 모드 5 (유닛 2 칸을 봄).
// [16번 수정 2026-11-09: 관리자 2(g_fbCtrlMode2)·모드 g_fbCmStdSched2 → 접속점 그룹 관리자 g_fbCtrlMode1·g_fbCmStdSched1의 유닛 2 칸] EMS 명령은 MQTT 수신 칸(GVL_MQTT.g_astPcsCommand[1] = PCS2)에 직접 넣음 (브로커 없이)
// A: 켠 직후 EMS P 없음 → 0 / B: 방전 100 → 100 / C: 충전 50 → -50 / D: 정지 → 0 (새 P 지령 대기)
// 조건이 2 s 이어지면 통과. 장비 쓰기(DEVICE_WRITE)와 무관하게 코어 고르기 결과(MAIN.fbSelect)까지 봄. 끝나면 모드 0, 운전 모드를 되돌림
VAR
	bStart		: BOOL;
	bDone		: BOOL;
	bPass		: BOOL;
	nStep		: UINT;
	wsStep		: WSTRING(80);
	wsFail		: WSTRING(80);
	(* 지금 값 *)
	nActive		: UINT;			// 접속점 그룹 관리자 켜진 모드 (5 = 스탠다드 스케줄)
	nModeState	: UINT;			// 모드 q_nState (0 = P 냄, 2 = EMS 끊김, 3 = 새 지령 대기)
	fModeP		: REAL;			// 모드가 받아 둔 P
	bEmsAlive	: BOOL;			// EMS 지령원 유효
	fMgrP		: REAL;			// 접속점 그룹 관리자 출력 (유닛 2 칸)
	bMgrP		: BOOL;
	stPick		: ST_Pick;		// 코어 고르기 결과 (Auto 유닛 2)
	(* 판정 *)
	bA			: BOOL;
	bB			: BOOL;
	bC			: BOOL;
	bD			: BOOL;
	fB			: REAL;
	fC			: REAL;
	(* 내부 *)
	nU2			: UINT := 2;
	eOpModeBak	: E_OpMode;
	bBackedUp	: BOOL;
	bCond		: BOOL;
	nLastStep	: UINT;
	tonStep		: TON;
	tonOk		: TON;
	stOut		: ST_SourceOutput;
END_VAR

// 지금 값
nActive		:= GVL_SITE.g_fbCtrlMode1.q_nActive;
stOut		:= GVL_SITE.g_fbCtrlMode1.Output;
IF nU2 >= 1 AND nU2 <= GVL_PARAM.UNIT_COUNT THEN
	nModeState	:= GVL_SITE.g_fbCmStdSched1.q_anState[nU2];
	fModeP		:= GVL_SITE.g_fbCmStdSched1.q_afPCmd[nU2];
	bEmsAlive	:= GVL_SITE.g_fbCmStdSched1.i_astCmd[nU2].bAlive;
	bMgrP	:= stOut.astUnit[nU2].bPSetActive;
	fMgrP	:= stOut.astUnit[nU2].fPSet;
	stPick	:= MAIN.fbSelect.q_astAutoUnitP[nU2];
END_IF

tonStep(IN := nStep >= 20 AND nStep < 900, PT := T#30S);
bCond := FALSE;

CASE nStep OF
	0:
		IF bStart THEN
			bStart := FALSE;	bDone := FALSE;	bPass := FALSE;	wsFail := "";
			bA := FALSE;	bB := FALSE;	bC := FALSE;	bD := FALSE;
			nStep := 10;
		ELSIF NOT bDone THEN
			wsStep := "대기: bStart := TRUE로 시작";
		END_IF

	10:	// PCS2 Auto
		wsStep := "PCS2 Auto 전환";
		IF nU2 > GVL_PARAM.UNIT_COUNT OR GVL_PARAM.PCS_COUNT < 2 THEN
			wsFail := "PCS·유닛이 2개 이상이어야 함";
			nStep := 900;
		ELSE
			eOpModeBak	:= GVL_PERSIST.g_aeOpMode[nU2];
			bBackedUp	:= TRUE;
			GVL_PERSIST.g_aeOpMode[nU2] := E_OpMode.Auto;
			nStep := 20;
		END_IF

	20:
		wsStep := "Auto 전환 대기";
		IF MAIN.fbModeSwitch.q_aeOpMode[nU2] = E_OpMode.Auto THEN
			GVL_SITE.g_fbCtrlMode1.i_nModeReq := 5;
			GVL_SITE.g_fbCtrlMode1.i_bRetry := TRUE;
			nStep := 30;
		END_IF

	30:
		wsStep := "스탠다드 스케줄 모드 켜는 중";
		IF nActive = 5 THEN
			nStep := 100;
		ELSIF GVL_SITE.g_fbCtrlMode1.q_eRefuse <> E_CtrlModeRefuse.None THEN
			wsFail := WCONCAT("모드 거부: ", GVL_SITE.g_fbCtrlMode1.M_ModeReasonText(i_nSlot := 5, i_nReason := GVL_SITE.g_fbCtrlMode1.q_nRefuseReason));
			nStep := 900;
		END_IF

	100: // A: 켠 직후, EMS P 없음 → 0
		wsStep := "A: EMS P 없음 → 0";
		bCond := nActive = 5 AND (nModeState = 3 OR nModeState = 2) AND bMgrP AND fMgrP = 0.0;
		IF tonOk.Q THEN
			bA := TRUE;
			M_Send(i_nType := 5, i_fValue := 100.0);		// 방전 100
			nStep := 110;
		END_IF
	110: // B: 방전 100
		wsStep := "B: EMS 방전 100 → 100";
		bCond := nModeState = 0 AND ABS(fModeP - 100.0) < 0.01 AND bMgrP AND ABS(fMgrP - 100.0) < 0.01
			AND stPick.bActive AND ABS(stPick.fValue - 100.0) < 0.01 AND stPick.nModule = GVL_SITE.g_fbCtrlMode1.ModuleId;
		IF tonOk.Q THEN
			bB := TRUE;	fB := stPick.fValue;
			M_Send(i_nType := 4, i_fValue := 50.0);		// 충전 50
			nStep := 120;
		END_IF
	120: // C: 충전 50
		wsStep := "C: EMS 충전 50 → -50";
		bCond := nModeState = 0 AND ABS(fMgrP + 50.0) < 0.01 AND stPick.bActive AND ABS(stPick.fValue + 50.0) < 0.01;
		IF tonOk.Q THEN
			bC := TRUE;	fC := stPick.fValue;
			M_Send(i_nType := 2, i_fValue := 0.0);		// 정지
			nStep := 130;
		END_IF
	130: // D: 정지 → 0 (새 P 지령 대기)
		wsStep := "D: EMS 정지 → 0";
		bCond := nModeState = 3 AND bMgrP AND fMgrP = 0.0 AND stPick.bActive AND stPick.fValue = 0.0;
		IF tonOk.Q THEN
			bD := TRUE;
			nStep := 900;
		END_IF

	900: // 정리
		GVL_SITE.g_fbCtrlMode1.i_nModeReq := 0;
		IF bBackedUp THEN
			GVL_PERSIST.g_aeOpMode[nU2] := eOpModeBak;
			bBackedUp := FALSE;
		END_IF
		bPass := bA AND bB AND bC AND bD AND wsFail = "";
		bDone := TRUE;
		IF bPass THEN
			wsStep := "끝: 통과";
		ELSE
			wsStep := "끝: 실패 (wsFail·구간 결과 확인)";
		END_IF
		nStep := 0;
END_CASE

tonOk(IN := bCond AND nStep = nLastStep, PT := T#2S);
IF tonStep.Q AND nStep >= 20 AND nStep < 900 THEN
	wsFail	:= WCONCAT("시간 초과: ", wsStep);
	nStep	:= 900;
END_IF
IF nStep <> nLastStep THEN
	tonStep(IN := FALSE);
	tonOk(IN := FALSE);
	nLastStep := nStep;
END_IF

METHOD PRIVATE M_Send		// EMS 명령 레코드 하나를 MQTT 수신 칸에 넣음 (PCS2 = 칸 1). 값을 먼저, 종류를 마지막에 (MqttTask가 종류를 보고 처리)
VAR_INPUT
	i_nType		: UDINT;	// PCS CommandType: 1 Run, 2 Stop, 3 Standby, 4 충전, 5 방전
	i_fValue	: REAL;		// kW
END_VAR
GVL_MQTT.g_astPcsCommand[1].DeviceIndex	:= 2;	// PCS2 (번호 1부터) [1부터 2026-11-10]
GVL_MQTT.g_astPcsCommand[1].Value		:= i_fValue;
GVL_MQTT.g_astPcsCommand[1].CommandType	:= i_nType;
END_METHOD

END_PROGRAM

// ---- 90_Project/PRG_Redundancy.TcPOU
PROGRAM PRG_Redundancy		// 이중화 태스크에서 부름 (높은 우선순위). 이 PLC의 역할(Primary/Secondary)과 지금 장비에 쓰는지(Active)를 GVL_IF에 씀
VAR
	fbGetNetId		: FB_GetLocalAmsNetID;	// 이 PLC의 AMS Net ID 읽기 (시작 때 한 번)
	sMyNetId		: T_AmsNetId;			// 읽은 이 PLC의 Net ID (온라인 확인용: RED_SET에 적을 값)
	bNetIdRead		: BOOL;					// Net ID를 읽었음
	tLastScan		: TIME;				// 지난 스캔의 시스템 시각 (멈췄다 이어짐 감지)
	bScanned		: BOOL;				// 첫 스캔을 지남 (시작 때는 이어짐으로 안 봄)
	bResume			: BOOL;				// 이번 스캔이 멈췄다 이어진 첫 스캔
	fbRedSync		: FB_RedSync;			// 운영 설정 동기화 (Active → Standby)
	fbRedState		: FB_RedState;			// 역할 + 상대 상태 → Active 판단
	fbRedLink		: FB_RedLink;			// 상대 PLC와 EAP 하트비트·접점 신호 (I/O는 이 인스턴스에 연결)
END_VAR

(* 0) 멈췄다 이어짐 감지: ADS·XAE의 Stop/Run은 변수를 초기화하지 않고 이어서 돎. 이전 스캔과 시스템 시각이 1 s 넘게 벌어지면 멈췄던 것으로 보고 상태를 Init부터 다시 정함 *)
bResume := bScanned AND (TIME() - tLastScan) > T#1S;
bScanned := TRUE;
tLastScan := TIME();
IF bResume AND GVL_SITE.RED_SET.bUse THEN
	GVL_IF.g_nRedResumeCount	:= GVL_IF.g_nRedResumeCount + 1;
	GVL_IF.g_bRedActive			:= FALSE;		// 옛 Active를 상대에게 알리거나 장비에 쓰지 않도록 이 스캔부터 내림
	GVL_IF.g_bRedWrite			:= FALSE;
	GVL_IF.g_eRedState			:= E_RedState.Init;
END_IF

(* 1) 역할: 이중화를 안 쓰면 Primary. 쓰면 이 PLC Net ID를 GVL_SITE.RED_SET과 비교 *)
IF NOT GVL_SITE.RED_SET.bUse THEN
	GVL_IF.g_eRedRole := E_RedRole.Primary;
ELSIF NOT bNetIdRead THEN
	GVL_IF.g_eRedRole := E_RedRole.Reading;
	fbGetNetId(bExecute := TRUE);
	IF NOT fbGetNetId.bBusy THEN
		IF NOT fbGetNetId.bError THEN
			sMyNetId	:= fbGetNetId.AddrString;
			bNetIdRead	:= TRUE;
		END_IF
		fbGetNetId(bExecute := FALSE);		// 오류면 다음 스캔에 다시 읽음
	END_IF
ELSIF sMyNetId = GVL_SITE.RED_SET.sPrimaryNetId THEN
	GVL_IF.g_eRedRole := E_RedRole.Primary;
ELSIF sMyNetId = GVL_SITE.RED_SET.sSecondaryNetId THEN
	GVL_IF.g_eRedRole := E_RedRole.Secondary;
ELSE
	GVL_IF.g_eRedRole := E_RedRole.NoMatch;		// 설정 오류 (FB_ConfigCheck)
END_IF

(* 2) 상대 PLC 상태: EAP 하트비트와 접점 신호를 보고 판정. 이중화를 안 쓰면 보내지도 않음. 내 Active는 지난 스캔 값을 보냄 *)
IF GVL_SITE.RED_SET.bUse THEN
	fbRedLink(	i_stSet	:= GVL_SITE.RED_SET,
				i_eRole	:= GVL_IF.g_eRedRole,
				i_bActive	:= GVL_IF.g_bRedActive,
				i_eState	:= GVL_IF.g_eRedState);
	GVL_IF.g_nRedSeq			:= fbRedLink.q_nTxCount;
	GVL_IF.g_ePeerState		:= fbRedLink.q_ePeer;
	GVL_IF.g_bPeerEapOk		:= fbRedLink.q_bEapOk;
	GVL_IF.g_bPeerWireOk		:= fbRedLink.q_bWireOk;
	GVL_IF.g_nPeerRole		:= fbRedLink.q_stPeer.nRole;
	GVL_IF.g_bPeerActive		:= fbRedLink.q_stPeer.bActive;
	GVL_IF.g_nPeerState		:= fbRedLink.q_stPeer.nState;
	GVL_IF.g_bPeerWireActive	:= fbRedLink.q_bPeerWireActive;
	GVL_IF.g_bRedRoleConflict	:= fbRedLink.q_bRoleConflict;
ELSE
	GVL_IF.g_ePeerState		:= E_RedPeer.Unknown;
	GVL_IF.g_bPeerEapOk		:= FALSE;
	GVL_IF.g_bPeerWireOk		:= FALSE;
	GVL_IF.g_bRedRoleConflict	:= FALSE;
	GVL_IF.g_nPeerState		:= 0;
END_IF

(* 3) 동기화: 운영 설정을 상대에게 보내고, 내가 Active가 아니고 상대가 Active이면 받은 값으로 맞춤
   동기화 대상 = GVL_PERSIST의 운영 설정 (재기동 기록·모듈 설정 묶음 제외) + 제어 모드 요청. 대상을 늘리면 ST_RedSyncCfg와 FB_RedSync의 보내기·맞추기에 추가 *)
IF GVL_SITE.RED_SET.bUse THEN
	fbRedSync(	i_bUse		:= TRUE,
				i_bApply	:= GVL_IF.g_eRedState <> E_RedState.Active AND GVL_IF.g_bPeerEapOk AND GVL_IF.g_bPeerActive);
	GVL_IF.g_bSyncInSync	:= fbRedSync.q_bInSync;
	GVL_IF.g_bSyncFresh		:= fbRedSync.q_bFresh;
	GVL_IF.g_nSyncApplied	:= fbRedSync.q_nApplied;
ELSE
	GVL_IF.g_bSyncInSync	:= FALSE;
	GVL_IF.g_bSyncFresh		:= FALSE;
END_IF

(* 4) Active: 역할과 상대 상태로 정함 (FB_RedState). 두 PLC가 동시에 Active가 되지 않음. Secondary 승격(절체)·Primary 복귀 포함 *)
fbRedState(	i_bUse			:= GVL_SITE.RED_SET.bUse,
			i_stSet			:= GVL_SITE.RED_SET,
			i_eRole			:= GVL_IF.g_eRedRole,
			i_ePeer			:= GVL_IF.g_ePeerState,
			i_bPeerActive	:= (GVL_IF.g_bPeerEapOk AND GVL_IF.g_bPeerActive) OR (GVL_IF.g_bPeerWireOk AND GVL_IF.g_bPeerWireActive),
			i_bPeerHandover	:= GVL_IF.g_bPeerEapOk AND GVL_IF.g_nPeerState = TO_INT(E_RedState.Handover),
			i_bRoleConflict	:= GVL_IF.g_bRedRoleConflict,
			i_bReset		:= bResume AND GVL_SITE.RED_SET.bUse,
			i_bSyncDone		:= GVL_IF.g_bSyncInSync);
GVL_IF.g_eRedState	:= fbRedState.q_eState;
GVL_IF.g_bRedActive	:= fbRedState.q_bActive;
GVL_IF.g_bRedWrite	:= fbRedState.q_bWrite;
GVL_IF.g_nRedSwitchCount	:= fbRedState.q_nSwitchCount;
GVL_IF.g_eRedSwitch	:= fbRedState.q_eLastSwitch;

END_PROGRAM

// ---- 10_Core/90_Redundancy/FB_RedSync.TcPOU
FUNCTION_BLOCK FB_RedSync		// 동기화: 이 PLC의 운영 설정(GVL_PERSIST, 모듈 설정 묶음 제외)과 제어 모드 요청(PCS마다)을 EAP로 매 스캔 상대에게 보내고, 상대가 Active이고 내가 Active가 아닐 때 받은 값으로 내 설정을 맞춘다
(* - 보내는 값은 EAP 변수 1개: 운영 설정(_stTx, ST_RedSyncCfg). 받는 값도 같은 모양(_stRx)
   - 모듈 설정 묶음(GVL_PERSIST.g_stModuleSet)은 동기화하지 않음: HMI가 두 PLC 모두에 씀 (PLC가 꺼져 있던 동안 바꾼 값은 복귀 전에 HMI에서 다시 쓸 것)
   - 맞추기: i_bApply일 때만, 값이 다른 것만 덮어씀 (같으면 안 씀: 저장을 불필요하게 만들지 않음). 바꾼 것이 없으면 q_bInSync
   - 살아 있음: _stRx.nSeq가 i_tTimeout 안에 바뀌어야 함 (q_bFresh)
   - 2026-11-23 UPS 항목 추가 (명세 RED-01 v2.43): UPS 설정 보관값·사고 대응 스위치. 형식 번호 2. BMS 랙 선택표는 동기화하지 않음 (실제 랙 상태로 씀)
   - 2026-11-25 사고 대응 된 동작 비트 추가 (명세 RED-01 v2.49): 보내고, 대기 쪽은 GVL_IF.g_awPeerRespDone에 기억만 함 (설정 아님: 일치·횟수에 안 넣음). 형식 번호 3
   - I/O(AT %I*·%Q)는 설치할 때 XAE에서 연결. 인스턴스는 RedundancyTask의 PRG_Redundancy에 둠. 두 PLC 프로그램이 같아야 함 *)
VAR_INPUT
	i_bUse			: BOOL;
	i_bApply		: BOOL;				// 받은 값을 내 설정에 덮어써도 됨 (내가 Active가 아니고 상대가 Active이며 통신 정상)
	i_tTimeout		: TIME := T#2S;		// 새 값이 이 시간 안에 안 오면 낡은 것
END_VAR
VAR_OUTPUT
	q_bInSync		: BOOL;				// 받은 값이 낡지 않았고 내 설정이 그와 같음 (i_bApply일 때만 TRUE)
	q_bFresh		: BOOL;				// 상대가 보낸 값이 낡지 않음
	q_nApplied		: UDINT;			// 받은 값으로 덮어쓴 횟수 (필드 단위)
END_VAR
VAR
	(* I/O: XAE에서 연결 *)
	_stTx			AT %Q* : ST_RedSyncCfg;
	_stRx			AT %I* : ST_RedSyncCfg;

	_nLastSeq		: UDINT;
	_tonFresh		: TON;
END_VAR
VAR_TEMP
	bNew			: BOOL;
	bEq				: BOOL;
END_VAR

IF NOT i_bUse THEN
	RETURN;
END_IF

(* 1) 보내기 *)
_stTx.nProtoVer	:= 4;	// 명세 RED-01 v2.51 (v2.49: 3)
_stTx.nSeq		:= _stTx.nSeq + 1;
_stTx.nModeReq1	:= GVL_SITE.g_fbCtrlMode1.i_nModeReq;
_stTx.aeOpMode := GVL_PERSIST.g_aeOpMode;
_stTx.astGroupSet := GVL_PERSIST.g_astGroupSet;
_stTx.astManualPolicy := GVL_PERSIST.g_astManualPolicy;
_stTx.astSourceReg := GVL_PERSIST.g_astSourceReg;
_stTx.astLimitReg := GVL_PERSIST.g_astLimitReg;
_stTx.astPermitReg := GVL_PERSIST.g_astPermitReg;
_stTx.astCompReg := GVL_PERSIST.g_astCompReg;
_stTx.astRuleCfg := GVL_PERSIST.g_astRuleCfg;
_stTx.astOutputCfg := GVL_PERSIST.g_astOutputCfg;
_stTx.astUnitRuleReg := GVL_PERSIST.g_astUnitRuleReg;
_stTx.astBatRuleReg := GVL_PERSIST.g_astBatRuleReg;
_stTx.stCmdFilter := GVL_PERSIST.g_stCmdFilter;
_stTx.stManualCmdSet := GVL_PERSIST.g_stManualCmdSet;
_stTx.stSeqSet := GVL_PERSIST.g_stSeqSet;
_stTx.stBrokerWatch := GVL_PERSIST.g_stBrokerWatch;	// [9번 수정 2026-11-09: 추가]
_stTx.astUpsDesired := GVL_PERSIST.g_astUpsDesired;	// 명세 RED-01 v2.43
_stTx.bUpsSafetyRespEnable := GVL_PERSIST.g_bUpsSafetyRespEnable;
_stTx.awUpsRespDone := GVL_IF.g_awUpsRespDone;	// 명세 RED-01 v2.49 (MAIN이 씀)

(* 2) 받기: 새 값이 오는지 *)
bNew := _stRx.nSeq <> _nLastSeq;
_nLastSeq := _stRx.nSeq;
_tonFresh(IN := NOT bNew, PT := i_tTimeout);
q_bFresh := _stRx.nProtoVer = 4 AND _stRx.nSeq <> 0 AND NOT _tonFresh.Q;

(* 3) 맞추기: 내가 Active가 아니고 상대가 Active일 때만 다른 것만 덮어씀 *)
q_bInSync := FALSE;
IF i_bApply AND q_bFresh THEN
	bEq := TRUE;
	IF GVL_SITE.g_fbCtrlMode1.i_nModeReq <> _stRx.nModeReq1 THEN
		GVL_SITE.g_fbCtrlMode1.i_nModeReq := _stRx.nModeReq1;
		q_nApplied := q_nApplied + 1;
		bEq := FALSE;
	END_IF
	IF MEMCMP(ADR(GVL_PERSIST.g_aeOpMode), ADR(_stRx.aeOpMode), SIZEOF(_stRx.aeOpMode)) <> 0 THEN
		GVL_PERSIST.g_aeOpMode := _stRx.aeOpMode;
		q_nApplied := q_nApplied + 1;
		bEq := FALSE;
	END_IF
	IF MEMCMP(ADR(GVL_PERSIST.g_astGroupSet), ADR(_stRx.astGroupSet), SIZEOF(_stRx.astGroupSet)) <> 0 THEN
		GVL_PERSIST.g_astGroupSet := _stRx.astGroupSet;
		q_nApplied := q_nApplied + 1;
		bEq := FALSE;
	END_IF
	IF MEMCMP(ADR(GVL_PERSIST.g_astManualPolicy), ADR(_stRx.astManualPolicy), SIZEOF(_stRx.astManualPolicy)) <> 0 THEN
		GVL_PERSIST.g_astManualPolicy := _stRx.astManualPolicy;
		q_nApplied := q_nApplied + 1;
		bEq := FALSE;
	END_IF
	IF MEMCMP(ADR(GVL_PERSIST.g_astSourceReg), ADR(_stRx.astSourceReg), SIZEOF(_stRx.astSourceReg)) <> 0 THEN
		GVL_PERSIST.g_astSourceReg := _stRx.astSourceReg;
		q_nApplied := q_nApplied + 1;
		bEq := FALSE;
	END_IF
	IF MEMCMP(ADR(GVL_PERSIST.g_astLimitReg), ADR(_stRx.astLimitReg), SIZEOF(_stRx.astLimitReg)) <> 0 THEN
		GVL_PERSIST.g_astLimitReg := _stRx.astLimitReg;
		q_nApplied := q_nApplied + 1;
		bEq := FALSE;
	END_IF
	IF MEMCMP(ADR(GVL_PERSIST.g_astPermitReg), ADR(_stRx.astPermitReg), SIZEOF(_stRx.astPermitReg)) <> 0 THEN
		GVL_PERSIST.g_astPermitReg := _stRx.astPermitReg;
		q_nApplied := q_nApplied + 1;
		bEq := FALSE;
	END_IF
	IF MEMCMP(ADR(GVL_PERSIST.g_astCompReg), ADR(_stRx.astCompReg), SIZEOF(_stRx.astCompReg)) <> 0 THEN
		GVL_PERSIST.g_astCompReg := _stRx.astCompReg;
		q_nApplied := q_nApplied + 1;
		bEq := FALSE;
	END_IF
	IF MEMCMP(ADR(GVL_PERSIST.g_astRuleCfg), ADR(_stRx.astRuleCfg), SIZEOF(_stRx.astRuleCfg)) <> 0 THEN
		GVL_PERSIST.g_astRuleCfg := _stRx.astRuleCfg;
		q_nApplied := q_nApplied + 1;
		bEq := FALSE;
	END_IF
	IF MEMCMP(ADR(GVL_PERSIST.g_astOutputCfg), ADR(_stRx.astOutputCfg), SIZEOF(_stRx.astOutputCfg)) <> 0 THEN
		GVL_PERSIST.g_astOutputCfg := _stRx.astOutputCfg;
		q_nApplied := q_nApplied + 1;
		bEq := FALSE;
	END_IF
	IF MEMCMP(ADR(GVL_PERSIST.g_astUnitRuleReg), ADR(_stRx.astUnitRuleReg), SIZEOF(_stRx.astUnitRuleReg)) <> 0 THEN
		GVL_PERSIST.g_astUnitRuleReg := _stRx.astUnitRuleReg;
		q_nApplied := q_nApplied + 1;
		bEq := FALSE;
	END_IF
	IF MEMCMP(ADR(GVL_PERSIST.g_astBatRuleReg), ADR(_stRx.astBatRuleReg), SIZEOF(_stRx.astBatRuleReg)) <> 0 THEN
		GVL_PERSIST.g_astBatRuleReg := _stRx.astBatRuleReg;
		q_nApplied := q_nApplied + 1;
		bEq := FALSE;
	END_IF
	IF MEMCMP(ADR(GVL_PERSIST.g_stCmdFilter), ADR(_stRx.stCmdFilter), SIZEOF(_stRx.stCmdFilter)) <> 0 THEN
		GVL_PERSIST.g_stCmdFilter := _stRx.stCmdFilter;
		q_nApplied := q_nApplied + 1;
		bEq := FALSE;
	END_IF
	IF MEMCMP(ADR(GVL_PERSIST.g_stManualCmdSet), ADR(_stRx.stManualCmdSet), SIZEOF(_stRx.stManualCmdSet)) <> 0 THEN
		GVL_PERSIST.g_stManualCmdSet := _stRx.stManualCmdSet;
		q_nApplied := q_nApplied + 1;
		bEq := FALSE;
	END_IF
	IF MEMCMP(ADR(GVL_PERSIST.g_stSeqSet), ADR(_stRx.stSeqSet), SIZEOF(_stRx.stSeqSet)) <> 0 THEN
		GVL_PERSIST.g_stSeqSet := _stRx.stSeqSet;
		q_nApplied := q_nApplied + 1;
		bEq := FALSE;
	END_IF
	IF MEMCMP(ADR(GVL_PERSIST.g_stBrokerWatch), ADR(_stRx.stBrokerWatch), SIZEOF(_stRx.stBrokerWatch)) <> 0 THEN	// [9번 수정 2026-11-09: 추가]
		GVL_PERSIST.g_stBrokerWatch := _stRx.stBrokerWatch;
		q_nApplied := q_nApplied + 1;
		bEq := FALSE;
	END_IF
	// UPS 항목 (명세 RED-01 v2.43)
	IF MEMCMP(ADR(GVL_PERSIST.g_astUpsDesired), ADR(_stRx.astUpsDesired), SIZEOF(_stRx.astUpsDesired)) <> 0 THEN
		GVL_PERSIST.g_astUpsDesired := _stRx.astUpsDesired;
		q_nApplied := q_nApplied + 1;
		bEq := FALSE;
	END_IF
	IF GVL_PERSIST.g_bUpsSafetyRespEnable <> _stRx.bUpsSafetyRespEnable THEN
		GVL_PERSIST.g_bUpsSafetyRespEnable := _stRx.bUpsSafetyRespEnable;
		q_nApplied := q_nApplied + 1;
		bEq := FALSE;
	END_IF
	q_bInSync := bEq;
	// 사고 대응 된 동작 (명세 RED-01 v2.49): 설정이 아니므로 기억만 함. 내가 Active가 되면 MAIN이 이어받음
	GVL_IF.g_awPeerRespDone := _stRx.awUpsRespDone;
END_IF

END_FUNCTION_BLOCK

// ---- 10_Core/90_Redundancy/FB_RedState.TcPOU
FUNCTION_BLOCK FB_RedState		// 이중화 상태 기계 (순수 로직). 역할 + 상대 상태 → 이 PLC가 Active인지, 장비에 써도 되는지. 두 PLC가 동시에 Active가 되지 않게 함
(* 규칙
   - 이중화를 안 쓰면 항상 Active이고 바로 쓴다
   - 역할 설정 오류(NoMatch) 또는 두 PLC 역할이 같음 → Failed (둘 다 장비에 쓰지 않음)
   - Primary: 시작하면 상대 상태를 볼 때까지 Init. 상대가 Active가 아니면 Active, 이미 Active이면 뺏지 않고 Standby
   - 절체: Secondary는 상대가 Lost(EAP·접점 둘 다 끊김)이고 tTakeoverDelay가 지나면 Active (Standby → Active)
   - 복귀: Primary가 Standby에서 상대(Secondary)가 Active이고 통신이 tFailbackStable 동안 정상이면 Handover(넘겨받기 요청)로 감.
     Secondary는 상대가 Handover이면 Active를 내려놓고 Standby로. Primary는 상대가 Active가 아니게 되면 Active.
     tHandoverTimeout 안에 안 내려놓으면 Primary가 Standby로 돌아가 다시 기다림. 둘 다 안 쓰는 틈이 생기지만 둘 다 쓰는 일은 없음
   - 둘 다 Active로 보이면 Secondary가 Standby로 물러남 (Primary 우선)
   - 상대 Active = EAP 하트비트의 Active (EAP 정상일 때) 또는 Active 접점 (접점 정상일 때)
   - PLC가 멈췄다 이어지면(i_bReset) Init부터 다시 정함: 멈춘 사이 상대가 Active를 넘겨받았을 수 있으므로 옛 Active를 이어 쓰지 않고, 상대 상태를 본 뒤 Standby로 들어가 복귀 절차를 밟음
   - 장비에 쓰는 허가(q_bWrite)는 Active가 된 뒤 tWriteHold가 지나야 켜짐 (승격 직후 계산이 안정되기를 기다림). Active가 아니게 되면 바로 꺼짐 *)
VAR_INPUT
	i_bUse			: BOOL;				// GVL_SITE.RED_SET.bUse
	i_stSet			: ST_RedSet;		// 시간 설정
	i_eRole			: E_RedRole;
	i_ePeer			: E_RedPeer;
	i_bPeerActive	: BOOL;				// 상대가 Active (EAP 또는 접점. 정상인 쪽만 반영해서 넘길 것)
	i_bPeerHandover	: BOOL;				// 상대가 Handover라고 알림 (EAP 정상일 때만)
	i_bRoleConflict	: BOOL;				// 두 PLC 역할이 같음 (FB_RedPeerMonitor)
	i_bReset		: BOOL;				// PLC가 멈췄다 이어짐: 상태를 Init부터 다시 정함 (멈춘 사이 상대가 Active를 넘겨받았을 수 있음)
	i_bSyncDone		: BOOL := TRUE;		// 복귀 전에 상대에게서 받을 값 동기화가 끝났음 (4단계에서 연결. 지금은 항상 TRUE)
END_VAR
VAR_OUTPUT
	q_eState		: E_RedState;
	q_bActive		: BOOL;				// Active 상태 (상대에게 알림)
	q_bWrite		: BOOL;				// 장비에 써도 됨 (Active + 쓰기 대기 지남)
	q_nSwitchCount	: UDINT;			// Active가 바뀐 횟수 (들어가거나 나옴)
	q_eLastSwitch	: E_RedSwitch;		// 마지막으로 바뀐 이유
END_VAR
VAR
	_ePrev			: E_RedState;
	_tonTakeover	: TON;
	_tonFailback	: TON;
	_tonHandover	: TON;
	_tonHold		: TON;
END_VAR

// 타이머는 매 스캔 부름
_tonTakeover(IN := i_eRole = E_RedRole.Secondary AND q_eState = E_RedState.Standby AND i_ePeer = E_RedPeer.Lost, PT := i_stSet.tTakeoverDelay);
_tonFailback(IN := i_eRole = E_RedRole.Primary AND q_eState = E_RedState.Standby AND i_ePeer = E_RedPeer.Alive AND i_bPeerActive AND i_bSyncDone, PT := i_stSet.tFailbackStable);
_tonHandover(IN := q_eState = E_RedState.Handover, PT := i_stSet.tHandoverTimeout);

IF i_bReset THEN
	q_eState := E_RedState.Init;
ELSIF NOT i_bUse THEN
	q_eState := E_RedState.Active;
ELSIF i_eRole = E_RedRole.NoMatch OR i_bRoleConflict THEN
	q_eState := E_RedState.Failed;
ELSIF i_eRole = E_RedRole.Reading THEN
	q_eState := E_RedState.Init;
ELSE
	IF q_eState = E_RedState.Failed THEN
		q_eState := E_RedState.Init;		// 오류가 풀리면 처음부터 다시 정함
	END_IF
	CASE q_eState OF
	E_RedState.Init:
		IF i_eRole = E_RedRole.Secondary THEN
			q_eState := E_RedState.Standby;
		ELSIF i_ePeer <> E_RedPeer.Unknown THEN		// Primary: 상대 상태를 본 뒤 정함
			IF i_bPeerActive THEN
				q_eState := E_RedState.Standby;
			ELSE
				q_eState := E_RedState.Active;
				q_eLastSwitch := E_RedSwitch.Start;
			END_IF
		END_IF
	E_RedState.Standby:
		IF i_eRole = E_RedRole.Secondary THEN
			IF _tonTakeover.Q THEN
				q_eState := E_RedState.Active;		// 절체
				q_eLastSwitch := E_RedSwitch.PeerLost;
			END_IF
		ELSIF i_ePeer <> E_RedPeer.Unknown THEN		// Primary
			IF NOT i_bPeerActive THEN
				q_eState := E_RedState.Active;		// 상대가 Active가 아님 (정지·대기)
				q_eLastSwitch := E_RedSwitch.Start;
			ELSIF _tonFailback.Q THEN
				q_eState := E_RedState.Handover;	// 복귀: 상대에게 Active를 내려놓으라고 알림
			END_IF
		END_IF
	E_RedState.Handover:
		IF NOT i_bPeerActive THEN
			q_eState := E_RedState.Active;			// 상대가 내려놓음 (또는 사라짐)
			q_eLastSwitch := E_RedSwitch.Failback;
		ELSIF _tonHandover.Q OR i_ePeer <> E_RedPeer.Alive THEN
			q_eState := E_RedState.Standby;			// 포기하고 처음부터 다시 기다림
		END_IF
	E_RedState.Active:
		IF i_eRole = E_RedRole.Secondary AND (i_bPeerActive OR i_bPeerHandover) THEN
			q_eState := E_RedState.Standby;			// Primary에 양보
			q_eLastSwitch := E_RedSwitch.Yield;
		END_IF
	ELSE
		q_eState := E_RedState.Init;
	END_CASE
END_IF

// Active가 들어가거나 나올 때 횟수
IF (q_eState = E_RedState.Active) <> (_ePrev = E_RedState.Active) THEN
	q_nSwitchCount := q_nSwitchCount + 1;
END_IF
_ePrev := q_eState;

q_bActive := q_eState = E_RedState.Active;
_tonHold(IN := q_bActive, PT := i_stSet.tWriteHold);
q_bWrite := q_bActive AND (_tonHold.Q OR NOT i_bUse);

END_FUNCTION_BLOCK

// ---- 10_Core/90_Redundancy/FB_RedLink.TcPOU
FUNCTION_BLOCK FB_RedLink		// 이중화 연결: EAP 하트비트 보내기·받기 + 접점 신호(EL2004 출력·EL1004 입력) 보내기·받기 + 상대 상태 판정 (FB_RedPeerMonitor)
(* - I/O 연결(AT %I*·%Q)은 설치할 때 XAE에서 한다. 인스턴스는 RedundancyTask를 도는 PRG_Redundancy에 둔다
   - EAP 보내기 _stTx → 상대가 받음, 받기 _stRx ← 상대가 보냄, Quality _nEapQuality: EAP 변수 연결 (값 = 마지막 갱신 뒤 지난 시간, 100 us 단위)
   - 접점: _bDoAlive(EL2004 채널 1)는 주기적으로 뒤집음 → 상대 _bDiPeerAlive(EL1004 채널 1). _bDoActive(채널 2)는 이 PLC가 Active인 동안 TRUE → 상대 _bDiPeerActive(채널 2)
   - 두 PLC에 같은 프로그램을 넣고, 두 PLC의 I/O 연결이 서로 마주 보게 한다 *)
VAR_INPUT
	i_stSet			: ST_RedSet;
	i_eRole			: E_RedRole;
	i_bActive		: BOOL;
	i_eState		: E_RedState;		// 이 PLC의 이중화 상태 (상대에게 알림)
END_VAR
VAR_OUTPUT
	q_ePeer			: E_RedPeer;		// 상대 상태
	q_bEapOk		: BOOL;
	q_bWireOk		: BOOL;
	q_stPeer		: ST_RedHeartbeat;	// 상대가 보낸 역할·Active (EAP 정상일 때만)
	q_bPeerWireActive: BOOL;			// 상대 Active 접점 (EAP와 따로 보는 값)
	q_bRoleConflict	: BOOL;				// 두 PLC 역할이 같음
	q_nTxCount		: UDINT;			// 보낸 하트비트 수
END_VAR
VAR CONSTANT
	PULSE_HALF		: TIME := T#100MS;	// alive 접점을 뒤집는 간격 (접점 타임아웃보다 충분히 짧게)
END_VAR
VAR
	(* I/O: XAE에서 연결 *)
	_stTx			AT %Q* : ST_RedHeartbeat;
	_stRx			AT %I* : ST_RedHeartbeat;
	_nEapQuality	AT %I* : UINT;		// EAP Subscriber의 Quality = 갱신 안 된 시간 (100 us 단위). tEapTimeout 이하면 정상
	_bDoAlive		AT %Q* : BOOL;		// EL2004 채널 1
	_bDoActive		AT %Q* : BOOL;		// EL2004 채널 2
	_bDiPeerAlive	AT %I* : BOOL;		// EL1004 채널 1
	_bDiPeerActive	AT %I* : BOOL;		// EL1004 채널 2

	_fbMon			: FB_RedPeerMonitor;
	_tonPulse		: TON;
END_VAR

(* 1) 보내기 *)
q_nTxCount			:= q_nTxCount + 1;
_stTx.nProtoVer		:= 2;
_stTx.nCounter		:= q_nTxCount;
_stTx.nRole			:= TO_INT(i_eRole);
_stTx.bActive		:= i_bActive;
_stTx.nState		:= TO_INT(i_eState);

_tonPulse(IN := NOT _tonPulse.Q, PT := PULSE_HALF);		// Q가 한 스캔 켜질 때마다 뒤집음
IF _tonPulse.Q THEN
	_bDoAlive := NOT _bDoAlive;
END_IF
_bDoActive			:= i_bActive;

(* 2) 받아서 판정 *)
_fbMon(	i_stRx			:= _stRx,
		i_nMyRole		:= TO_INT(i_eRole),
		i_bEapQualityOk	:= UINT_TO_UDINT(_nEapQuality) <= TIME_TO_UDINT(i_stSet.tEapTimeout) * 10,	// Quality = 갱신 안 된 시간 (100 us 단위)
		i_bWireAlive	:= _bDiPeerAlive,
		i_tEapTimeout	:= i_stSet.tEapTimeout,
		i_tWireTimeout	:= i_stSet.tWireTimeout,
		i_tStartGrace	:= i_stSet.tStartGrace);
q_ePeer				:= _fbMon.q_ePeer;
q_bEapOk			:= _fbMon.q_bEapOk;
q_bWireOk			:= _fbMon.q_bWireOk;
q_stPeer			:= _fbMon.q_stPeer;
q_bPeerWireActive	:= _bDiPeerActive;
q_bRoleConflict		:= _fbMon.q_bRoleConflict;

END_FUNCTION_BLOCK

// ---- 10_Core/90_Redundancy/FB_RedPeerMonitor.TcPOU
FUNCTION_BLOCK FB_RedPeerMonitor		// 상대 PLC 상태 판정 (순수 로직: I/O를 직접 안 봄). EAP 하트비트(카운터가 바뀌고 Quality 정상)와 접점 신호(값이 바뀜)를 따로 보고 합침
// 판정 규칙: 둘 다 정상 = Alive, 한쪽만 끊김 = 그 통신 고장 (상대는 살아 있음, 절체 안 함), 둘 다 끊김 = Lost (절체 조건)
VAR_INPUT
	i_stRx			: ST_RedHeartbeat;	// 받은 EAP 하트비트
	i_bEapQualityOk	: BOOL;				// EAP Quality가 정상
	i_nMyRole		: INT;				// 이 PLC의 역할 (E_RedRole). 받은 역할이 같으면 내 프레임이 되돌아온 것으로 보고 무시
	i_bWireAlive	: BOOL;				// 상대 alive 접점(DI)의 지금 값. 상대가 주기적으로 뒤집음
	i_tEapTimeout	: TIME := T#500MS;	// 카운터가 이 시간 안 바뀌면 EAP 끊김
	i_tWireTimeout	: TIME := T#500MS;	// 접점이 이 시간 안 바뀌면 접점 끊김
	i_tStartGrace	: TIME := T#3S;		// 시작 직후 대기: 이 안에는 아직 못 봐도 Unknown
END_VAR
VAR_OUTPUT
	q_ePeer			: E_RedPeer;
	q_bEapOk		: BOOL;				// EAP 하트비트 정상
	q_bWireOk		: BOOL;				// 접점 신호 정상
	q_stPeer		: ST_RedHeartbeat;	// 상대가 보낸 값. EAP가 정상일 때만 채움 (아니면 0)
	q_bRoleConflict	: BOOL;				// 상대가 나와 같은 역할로 살아 있음 (두 PLC 역할 설정 오류). 접점도 살아 있을 때만 (내 프레임이 되돌아온 경우와 구분)
END_VAR
VAR
	_bInit			: BOOL;
	_nLastCount		: UDINT;
	_bLastWire		: BOOL;
	_bEapSeen		: BOOL;			// 시작 뒤 카운터가 바뀌는 것을 한 번이라도 봄
	_bWireSeen		: BOOL;
	_bSameSeen		: BOOL;
	_tonSame		: TON;
	_tonEap			: TON;
	_tonWire		: TON;
	_tonStart		: TON;
END_VAR
VAR_TEMP
	bEapMoved		: BOOL;
	bFromSelf		: BOOL;
	bSameMoved		: BOOL;
	bCntMoved		: BOOL;
	bWireMoved		: BOOL;
	stZero			: ST_RedHeartbeat;
END_VAR

IF NOT _bInit THEN
	_nLastCount	:= i_stRx.nCounter;
	_bLastWire	:= i_bWireAlive;
	_bInit		:= TRUE;
END_IF

// EAP: 카운터가 바뀌었고 Quality 정상이면 살아 있음. 안 바뀌는 시간이 길면 끊김 (상대 PLC가 멈추면 마지막 값이 그대로 남으므로 Quality만으로는 못 잡음)
bFromSelf		:= i_stRx.nRole = i_nMyRole;	// 상대와 내 역할은 항상 다름. 같으면 루프로 되돌아온 내 프레임 (또는 역할 설정 오류)
bCntMoved		:= i_bEapQualityOk AND i_stRx.nCounter <> _nLastCount;
bEapMoved		:= bCntMoved AND NOT bFromSelf;
_nLastCount		:= i_stRx.nCounter;
IF bEapMoved THEN
	_bEapSeen := TRUE;
END_IF
// 같은 역할 프레임이 계속 오는지 (Primary·Secondary일 때만. 시작 중 Reading끼리는 제외)
bSameMoved		:= bCntMoved AND bFromSelf AND (i_nMyRole = 1 OR i_nMyRole = 2);
IF bSameMoved THEN
	_bSameSeen := TRUE;
END_IF
_tonSame(IN := NOT bSameMoved, PT := i_tEapTimeout);
_tonEap(IN := NOT bEapMoved, PT := i_tEapTimeout);
q_bEapOk		:= _bEapSeen AND NOT _tonEap.Q AND i_bEapQualityOk AND NOT bFromSelf;

// 접점: 값이 바뀌면 살아 있음
bWireMoved		:= i_bWireAlive <> _bLastWire;
_bLastWire		:= i_bWireAlive;
IF bWireMoved THEN
	_bWireSeen := TRUE;
END_IF
_tonWire(IN := NOT bWireMoved, PT := i_tWireTimeout);
q_bWireOk		:= _bWireSeen AND NOT _tonWire.Q;
q_bRoleConflict	:= _bSameSeen AND NOT _tonSame.Q AND q_bWireOk;

_tonStart(IN := TRUE, PT := i_tStartGrace);

IF q_bEapOk AND q_bWireOk THEN
	q_ePeer := E_RedPeer.Alive;
ELSIF q_bWireOk THEN
	q_ePeer := E_RedPeer.EapLost;
ELSIF q_bEapOk THEN
	q_ePeer := E_RedPeer.WireLost;
ELSIF NOT _bEapSeen AND NOT _bWireSeen AND NOT _tonStart.Q THEN
	q_ePeer := E_RedPeer.Unknown;
ELSE
	q_ePeer := E_RedPeer.Lost;
END_IF

IF q_bEapOk THEN
	q_stPeer := i_stRx;
ELSE
	q_stPeer := stZero;
END_IF

END_FUNCTION_BLOCK

// ---- 20_Module/Common/FB_AuxIo.TcPOU
FUNCTION_BLOCK FB_AuxIo EXTENDS FB_DeviceBase IMPLEMENTS I_AuxDevice		// 벡호프 단자 I/O (EL1xxx 입력, EL2xxx 출력, EL3xxx 아날로그 입력, EL4xxx 아날로그 출력)
(* 점은 TwinCAT 화면에서 _abDi·_abDo·_anAi·_anAo 칸에 하나씩 연결. 점 번호 = 배열 칸 번호
   이 FB를 PlcTask가 아닌 태스크에서 쓰면 그 태스크 PRG 안에 선언 (GVL에 두면 TcContextName 필요) *)
VAR_INPUT
	i_afAiGain		: ARRAY[1..GVL_PARAM.AUX_AI_MAX] OF REAL;		// 아날로그 입력 = 원시값 × 배율 + 오프셋. 배율 0 = 1 (예: PT100 EL3202는 0.1)
	i_afAiOffset	: ARRAY[1..GVL_PARAM.AUX_AI_MAX] OF REAL;
	i_afAoGain		: ARRAY[1..GVL_PARAM.AUX_AO_MAX] OF REAL;		// 아날로그 출력 원시값 = 값 / 배율. 배율 0 = 1
END_VAR
VAR
	_abDi	AT %I*	: ARRAY[1..GVL_PARAM.AUX_DI_MAX] OF BOOL;
	_abDo	AT %Q*	: ARRAY[1..GVL_PARAM.AUX_DO_MAX] OF BOOL;
	_anAi	AT %I*	: ARRAY[1..GVL_PARAM.AUX_AI_MAX] OF INT;
	_anAo	AT %Q*	: ARRAY[1..GVL_PARAM.AUX_AO_MAX] OF INT;
	_bWcError AT %I* : BOOL;		// (선택) EtherCAT WcState 연결. 안 연결하면 늘 정상
END_VAR

METHOD M_Cycle
IF NOT _bWcError THEN
	M_MarkAlive();
END_IF
M_UpdateComm();
END_METHOD

PROPERTY Comm : BOOL
GET
Comm := _bComm;
END_GET
END_PROPERTY

METHOD M_GetBit : BOOL
VAR_INPUT
	i_nPoint	: UINT;
END_VAR
IF i_nPoint >= 1 AND i_nPoint <= GVL_PARAM.AUX_DI_MAX THEN
	M_GetBit := _abDi[i_nPoint];
END_IF
END_METHOD

METHOD M_GetValue : ST_Val
VAR_INPUT
	i_nPoint	: UINT;
END_VAR
IF i_nPoint >= 1 AND i_nPoint <= GVL_PARAM.AUX_AI_MAX THEN
	M_GetValue.fValue := INT_TO_REAL(_anAi[i_nPoint]) * SEL(i_afAiGain[i_nPoint] = 0, i_afAiGain[i_nPoint], 1.0) + i_afAiOffset[i_nPoint];
	M_GetValue.bValid := _bComm;
END_IF
END_METHOD

METHOD M_SetBit
VAR_INPUT
	i_nPoint	: UINT;
	i_bValue	: BOOL;
END_VAR
IF i_nPoint >= 1 AND i_nPoint <= GVL_PARAM.AUX_DO_MAX THEN
	_abDo[i_nPoint] := i_bValue;
END_IF
END_METHOD

METHOD M_SetValue
VAR_INPUT
	i_nPoint	: UINT;
	i_fValue	: REAL;
END_VAR
IF i_nPoint >= 1 AND i_nPoint <= GVL_PARAM.AUX_AO_MAX THEN
	// [결함 13 수정 2026-11-04: 값·게인이 숫자가 아니면 0 (LIMIT·REAL_TO_INT에서 FPU 예외). 원래 아래 줄만]
	IF F_RealOk(i_fValue) AND F_RealOk(i_afAoGain[i_nPoint]) THEN
		_anAo[i_nPoint] := REAL_TO_INT(LIMIT(-32768.0, i_fValue / SEL(i_afAoGain[i_nPoint] = 0, i_afAoGain[i_nPoint], 1.0), 32767.0));
	ELSE
		_anAo[i_nPoint] := 0;
	END_IF
END_IF
END_METHOD

END_FUNCTION_BLOCK

// ---- 10_Core/03_Base/FB_DeviceBase.TcPOU
FUNCTION_BLOCK ABSTRACT FB_DeviceBase EXTENDS FB_ModuleBase
VAR_INPUT
	i_tCommTimeout		: TIME := T#10S;	// 이 시간 동안 정상 응답이 없으면 통신 이상
	i_tReadPeriod		: TIME := T#200MS;	// 읽기 주기. 장비마다 GVL_SITE 인스턴스 선언에서 바꿈 (i_tCommTimeout보다 짧게)
END_VAR
VAR
	_bComm				: BOOL;		// 통신 정상
	_bAlive				: BOOL;		// 이번 스캔에 정상 응답(또는 하트비트 변화)이 있었음
	_bEverAlive			: BOOL;		// 부팅 후 한 번이라도 응답이 있었음
	_tonCommLoss		: TON;
	_fbRead				: FB_ReadTimer;
	_nWriteFails		: UINT;		// 잇달아 실패한 쓰기 수
	_bWriteFail			: BOOL;		// 쓰기 실패 (드라이버가 상태 bWriteFail에 넣음)
END_VAR
VAR CONSTANT
	WRITE_FAIL_COUNT	: UINT := 3;	// 쓰기가 이만큼 잇달아 실패하면 쓰기 실패로 봄 (한 번 성공하면 풀림)
END_VAR

METHOD PROTECTED M_MarkAlive
_bAlive		:= TRUE;
_bEverAlive	:= TRUE;
END_METHOD

METHOD PROTECTED M_IsReadTime : BOOL		// 읽을 때가 되면 TRUE (i_tReadPeriod마다). 스캔당 한 번만 부를 것
_fbRead(i_tPeriod := i_tReadPeriod);
M_IsReadTime := _fbRead.q_bDue;
END_METHOD

METHOD PROTECTED M_UpdateComm
// 마지막 정상 응답 이후 i_tCommTimeout이 지나면 통신 이상
_tonCommLoss(IN := NOT _bAlive, PT := i_tCommTimeout);
_bComm	:= _bEverAlive AND NOT _tonCommLoss.Q;	// 한 번도 응답이 없으면 정상으로 보지 않는다
_bAlive	:= FALSE;								// 다음 스캔을 위해 초기화
END_METHOD

METHOD PROTECTED M_MarkWriteResult		// 쓰기 결과를 알림 (드라이버가 쓰기 응답을 받을 때마다). 잇달아 WRITE_FAIL_COUNT번 실패하면 _bWriteFail, 한 번 성공하면 풀림
VAR_INPUT
	i_bOk	: BOOL;
END_VAR
IF i_bOk THEN
	_nWriteFails	:= 0;
	_bWriteFail		:= FALSE;
ELSE
	IF _nWriteFails < WRITE_FAIL_COUNT THEN
		_nWriteFails := _nWriteFails + 1;
	END_IF
	_bWriteFail := _nWriteFails >= WRITE_FAIL_COUNT;
END_IF
END_METHOD

END_FUNCTION_BLOCK

// ---- 10_Core/02_Util/FB_ReadTimer.TcPOU
FUNCTION_BLOCK FB_ReadTimer		// 읽기 주기 타이머: 읽을 때가 되면 그 스캔만 q_bDue = TRUE. 처음 호출 때 바로 TRUE
VAR_INPUT
	i_tPeriod		: TIME := T#200MS;	// 읽기 주기. T#0S면 매 스캔
END_VAR
VAR_OUTPUT
	q_bDue			: BOOL;
END_VAR
VAR
	_bStarted		: BOOL;
	_tonWait		: TON;
END_VAR

// 스캔당 한 번만 호출할 것
_tonWait(IN := _bStarted, PT := i_tPeriod);
q_bDue := NOT _bStarted OR _tonWait.Q;

IF q_bDue THEN
	_bStarted := TRUE;
	_tonWait(IN := FALSE, PT := i_tPeriod);	// 이번 스캔부터 다시 셈
	_tonWait(IN := TRUE, PT := i_tPeriod);
END_IF

END_FUNCTION_BLOCK

// ---- 20_Module/Mqtt/FB_SrcEms.TcPOU
FUNCTION_BLOCK FB_SrcEms EXTENDS FB_SourceBase		// 지령원: EMS (상위 플랫폼, MQTT command). 명령 핸들러(FB_EmsCommand)가 해석한 명령을 요청으로 냄
(* - 입력 i_stCmd는 MAIN(A_PassEmsCmd)이 GVL_IF에서 일관되게 복사해 넘긴다. 이 FB는 GVL을 보지 않는다
   - 상태 명령(PCS Run·Standby·Stop·EStop·Reset, 배터리 Close·Open): 번호가 바뀌면 새 명령. 큐에 넣고 스캔마다 1개씩 요청으로 낸다.
     받는 운전 모드는 등록표 stStateMode가 정한다. 배터리 Reset은 운전자 리셋(PCS Reset, 전체)으로 낸다
   - 충전·방전 P 지령: PCS 한 대의 kW를 그 PCS의 유닛들에 정격 비율로 나눠 유닛 지령(astUnit)으로 낸다.
     i_bPEnable이 TRUE일 때만 낸다 (기본 FALSE). 제어 모드(FB_CtrlModeMgr)와 어떻게 묶을지는 정해지면 여기서 연결 (상태 명령은 이 값과 무관하게 받음)
   - 새 메시지(nRxCount)나 새 명령이 만료 시간(등록 tExpire) 안에 오면 살아 있음. 끊기면 P 지령·요청 큐를 버린다 (돌아와도 옛 지령이 되살아나지 않음)
   - PMS가 켜진 뒤 처음 복사본은 번호만 맞춘다 (재기동 때 지난 명령을 실행하지 않음)
   - 배터리 비상정지(EStop)는 지령원 요청 종류에 없어 받지 않고 q_nUnsupported로 센다 *)
VAR_INPUT
	i_stCmd			: ST_IfEmsCmd;	// MAIN이 GVL_IF에서 복사한 명령 칸
	i_bValid		: BOOL;			// i_stCmd가 한 번이라도 일관되게 복사됨
	i_astUnitCfg	: ARRAY[1..GVL_PARAM.UNIT_COUNT] OF ST_UnitCfg;	// 유닛 ← PCS 번호 (명령은 PCS 번호로 옴)
	i_astBmsCfg		: ARRAY[1..GVL_PARAM.BMS_COUNT] OF ST_BmsCfg;	// BMS → 배터리 그룹
	i_bPEnable		: BOOL;			// 충전·방전 P 지령을 낼지 (기본 FALSE. 제어 모드와의 연결 방식이 정해질 때까지 끔)
END_VAR
VAR_OUTPUT
	q_nUnsupported	: UDINT;		// 받을 수 없는 명령 수 (배터리 비상정지)
	q_nQueueDrop	: UDINT;		// 큐가 가득 차 버린 요청 수
END_VAR
VAR CONSTANT
	QUEUE_PCS		: UINT := 16;
	QUEUE_BAT		: UINT := 8;
END_VAR
VAR
	_bSynced		: BOOL;
	_nRxCount		: UDINT;
	_anPcsSeq		: ARRAY[1..GVL_PARAM.PCS_COUNT] OF UDINT;
	_anPSeq			: ARRAY[1..GVL_PARAM.PCS_COUNT] OF UDINT;
	_anBatSeq		: ARRAY[1..GVL_PARAM.BMS_COUNT] OF UDINT;
	_abUnitP		: ARRAY[1..GVL_PARAM.UNIT_COUNT] OF BOOL;	// 이 유닛에 받아 둔 P 지령 있음
	_afUnitP		: ARRAY[1..GVL_PARAM.UNIT_COUNT] OF REAL;	// kW, 유닛 출력 (방전 +)
	_astPcsQ		: ARRAY[1..QUEUE_PCS] OF ST_PcsReq;
	_nPcsHead		: UINT := 1;
	_nPcsCount		: UINT;
	_astBatQ		: ARRAY[1..QUEUE_BAT] OF ST_BatReq;
	_nBatHead		: UINT := 1;
	_nBatCount		: UINT;
END_VAR

METHOD PRIVATE M_PushBat
VAR_INPUT
	i_eCmd		: E_BatCmd;
	i_nBatGroup	: UINT;
END_VAR
VAR
	nTail		: UINT;
END_VAR
IF _nBatCount >= QUEUE_BAT THEN
	q_nQueueDrop := q_nQueueDrop + 1;
	RETURN;
END_IF
nTail := ((_nBatHead + _nBatCount - 1) MOD QUEUE_BAT) + 1;
_astBatQ[nTail].eCmd		:= i_eCmd;
_astBatQ[nTail].nBatGroup	:= i_nBatGroup;
_nBatCount := _nBatCount + 1;
END_METHOD

METHOD PRIVATE M_PushPcs
VAR_INPUT
	i_eCmd		: E_PcsCmd;
	i_nUnit		: UINT;		// 0 = 그룹 전체
END_VAR
VAR
	nTail		: UINT;
END_VAR
IF _nPcsCount >= QUEUE_PCS THEN
	q_nQueueDrop := q_nQueueDrop + 1;
	RETURN;
END_IF
nTail := ((_nPcsHead + _nPcsCount - 1) MOD QUEUE_PCS) + 1;
_astPcsQ[nTail].eCmd	:= i_eCmd;
_astPcsQ[nTail].nUnit	:= i_nUnit;
_nPcsCount := _nPcsCount + 1;
END_METHOD

METHOD M_ReasonText : WSTRING(63)
VAR_INPUT
	i_nReason	: UINT;
END_VAR
M_ReasonText := "EMS 지령";
END_METHOD

METHOD M_UpdateOutput : BOOL
VAR
	p			: UINT;
	u			: UINT;
	b			: UINT;
	bFresh		: BOOL;
	bNewP		: BOOL;
	bAlgoOn		: BOOL;
	fSum		: REAL;
END_VAR
M_UpdateOutput := FALSE;

// 복사본이 아직 한 번도 없으면 기다림. 처음 받은 복사본은 번호만 맞춤 (지난 명령을 실행하지 않음)
IF NOT i_bValid THEN
	RETURN;
END_IF
IF NOT _bSynced THEN
	_bSynced := TRUE;
	_nRxCount := i_stCmd.nRxCount;
	FOR p := 1 TO GVL_PARAM.PCS_COUNT DO
		_anPcsSeq[p]	:= i_stCmd.astPcs[p].nSeq;
		_anPSeq[p]		:= i_stCmd.anPcsPSeq[p];
	END_FOR
	FOR b := 1 TO GVL_PARAM.BMS_COUNT DO
		_anBatSeq[b]	:= i_stCmd.astBat[b].nSeq;
	END_FOR
	RETURN;
END_IF

// 끊긴 상태(지난 스캔 기준)면 받아 둔 P 지령과 큐를 버림
IF _tonExpire.Q THEN
	FOR u := 1 TO GVL_PARAM.UNIT_COUNT DO
		_abUnitP[u] := FALSE;
	END_FOR
	_nPcsCount := 0;
	_nBatCount := 0;
END_IF

bFresh := FALSE;
bNewP := FALSE;
IF i_stCmd.nRxCount <> _nRxCount THEN
	_nRxCount := i_stCmd.nRxCount;
	bFresh := TRUE;
END_IF

// PCS: 상태 명령 → 그 PCS의 유닛마다 요청 (리셋은 전체 한 번), P 지령 → 유닛에 정격 비율로 나눔
FOR p := 1 TO GVL_PARAM.PCS_COUNT DO
	IF i_stCmd.astPcs[p].nSeq <> _anPcsSeq[p] THEN
		_anPcsSeq[p] := i_stCmd.astPcs[p].nSeq;
		bFresh := TRUE;
		IF i_stCmd.astPcs[p].eCmd = E_PcsCmd.Reset THEN
			M_PushPcs(E_PcsCmd.Reset, 0);
		ELSIF i_stCmd.astPcs[p].eCmd <> E_PcsCmd.None THEN
			FOR u := 1 TO GVL_PARAM.UNIT_COUNT DO
				IF i_astUnitCfg[u].nPcs = p THEN
					M_PushPcs(i_stCmd.astPcs[p].eCmd, u);
				END_IF
			END_FOR
		END_IF
	END_IF
	IF i_stCmd.anPcsPSeq[p] <> _anPSeq[p] THEN
		_anPSeq[p] := i_stCmd.anPcsPSeq[p];
		bFresh := TRUE;
		bNewP := TRUE;
		fSum := 0.0;
		FOR u := 1 TO GVL_PARAM.UNIT_COUNT DO
			IF i_astUnitCfg[u].nPcs = p THEN
				fSum := fSum + i_astUnitCfg[u].fPRated;
			END_IF
		END_FOR
		FOR u := 1 TO GVL_PARAM.UNIT_COUNT DO
			IF i_astUnitCfg[u].nPcs = p THEN
				_abUnitP[u] := TRUE;
				IF fSum > 0.0 THEN
					_afUnitP[u] := i_stCmd.afPcsP[p] * i_astUnitCfg[u].fPRated / fSum;
				ELSE
					_afUnitP[u] := 0.0;
				END_IF
			END_IF
		END_FOR
	END_IF
END_FOR

// BMS: 투입·개방은 배터리 그룹 요청, 리셋은 운전자 리셋
FOR b := 1 TO GVL_PARAM.BMS_COUNT DO
	IF i_stCmd.astBat[b].nSeq <> _anBatSeq[b] THEN
		_anBatSeq[b] := i_stCmd.astBat[b].nSeq;
		bFresh := TRUE;
		IF i_stCmd.astBat[b].eCmd = E_BatCmd.Close OR i_stCmd.astBat[b].eCmd = E_BatCmd.Open THEN
			M_PushBat(i_stCmd.astBat[b].eCmd, i_astBmsCfg[b].nBatGroup);
		ELSIF i_stCmd.astBat[b].eCmd = E_BatCmd.Reset THEN
			M_PushPcs(E_PcsCmd.Reset, 0);
		ELSE
			q_nUnsupported := q_nUnsupported + 1;
		END_IF
	END_IF
END_FOR

// 큐에서 한 스캔에 하나씩 요청으로 냄
IF _nPcsCount > 0 THEN
	_stOut.stPcsReq := _astPcsQ[_nPcsHead];
	_nPcsHead := (_nPcsHead MOD QUEUE_PCS) + 1;
	_nPcsCount := _nPcsCount - 1;
END_IF
IF _nBatCount > 0 THEN
	_stOut.stBatReq := _astBatQ[_nBatHead];
	_nBatHead := (_nBatHead MOD QUEUE_BAT) + 1;
	_nBatCount := _nBatCount - 1;
END_IF

// P 지령: 알고리즘이 선택된 그룹에서만. 받은 값은 새 명령이 올 때까지 유지 (만료되면 위에서 버림)
bAlgoOn := i_bPEnable;		// 등록 사용 여부(bEnable)는 FB_SourceBase가 처리 (꺼져 있으면 전부 지움)
FOR u := 1 TO GVL_PARAM.UNIT_COUNT DO
	_stOut.astUnit[u].bPSetActive	:= _abUnitP[u] AND bAlgoOn;
	_stOut.astUnit[u].fPSet			:= _afUnitP[u];
	_stOut.astUnit[u].bQSetActive	:= FALSE;
END_FOR
_stOut.bNewSet := bNewP AND bAlgoOn;

M_UpdateOutput := bFresh;
END_METHOD

END_FUNCTION_BLOCK

// ---- 20_Module/Driver/Plaspo/FB_PlaspoPcs.TcPOU
FUNCTION_BLOCK FB_PlaspoPcs EXTENDS FB_DeviceBase IMPLEMENTS I_Pcs		// 플라스포 PCS (Modbus TCP, 유닛 1개). 레지스터 맵은 Helios FB_PlaspoPcs와 같음
(* ---------------------------------------------------------------
   상태 (읽기 맵 → ST_UnitState)
   - 고장 비트 → Fault, 인버터 정지 → Stop
   - 운전 중이면서 마지막 상태 명령이 Standby → Standby, 그 밖의 운전 중 → Run
     (플라스포에는 Standby 상태가 따로 없어서 "운전 중 + 대기 모드(103 = 0)"를 Standby로 봄)
   명령 (레지스터: 값)
   - 기동    101: 55, 105: 1       - 정지·비상정지 101: 99, 105: 1 (비상정지 명령이 따로 없음)
   - 리셋    102: 33, 105: 1       - Standby  (정지 중이면 기동 먼저) 106: 1, 103: 0, 107: 0
   - 출력    P > 0 방전 103: 2, P < 0 충전 103: 1, 107: |P| × i_fPScale. 방향이 같으면 107만 씀
   - Q 지령은 이 맵에 없음 → 무시
   쓰기: 한 번에 레지스터 하나, 사이 간격 i_tWriteGap. 상태 명령이 출력보다 먼저.
         출력은 가장 최근 값만 보냄 (밀려 있으면 덮어씀)
   현장 확인: 유효전력 부호(i_bPInvert), 출력 레지스터 단위(i_fPScale)
   --------------------------------------------------------------- *)
VAR_INPUT
	i_sIpAddr		: STRING(15);
	i_nPort			: UINT := 502;
	i_nUnitId		: BYTE := 1;
	i_fPScale		: REAL := 1.0;		// 출력 레지스터(107) = kW × 배율
	i_bPInvert		: BOOL := TRUE;		// 읽은 유효전력 부호 뒤집기 (Helios: -acActive → 방전 +)
	i_tWriteGap		: TIME := T#300MS;	// 레지스터 쓰기 사이 간격 (Helios 300 ms)
	i_tTimeout		: TIME := T#1S;
END_VAR
VAR
	(* 읽기 *)
	_fbMbRead			: FB_MBReadRegs;
	_stReadMap			: ST_PlaspoPcsRaw;
	_bReadDue		: BOOL;
	_bReading		: BOOL;
	_bReadError		: BOOL;
	_nReadErrId		: UDINT;
	_stUnit			: ST_UnitState;
	_bStandbyMode	: BOOL;				// 마지막 상태 명령이 Standby
	(* 보낼 목록 (대기): 상태 명령은 가장 최근 것만, 출력은 가장 최근 값만 *)
	_anCmdRegAddr		: ARRAY[1..5] OF UINT;	// 보낼 상태 명령 (가장 최근 것만)
	_anCmdRegValue		: ARRAY[1..5] OF INT;
	_nCmdRegCount		: UINT;				// 0 = 없음
	_bPowerPending	: BOOL;
	_nPowerDir		: INT;				// 보낼 방향 (103 값): 0 그대로, 1 충전, 2 방전
	_nPowerAbs	: INT;				// 107
	_nDirWritten	: INT;				// 마지막으로 쓴 103
	(* 지금 보내는 목록 *)
	_fbMbWrite		: FB_MBWriteRegs;
	_anSendAddr		: ARRAY[1..5] OF UINT;
	_anSendValue		: ARRAY[1..5] OF INT;
	_nSendCount		: UINT;
	_nSendIdx		: UINT;
	_nWriteStep		: UINT;				// 0 다음 일 고르기, 1 쓰기 시작, 2 끝나기 기다림, 3 간격
	_bWriteError	: BOOL;
	_nWriteErrId	: UDINT;
	_tonWriteGap			: TON;
	_nCopyIdx			: UINT;				// 액션에서 쓰는 반복 변수
END_VAR

ACTION A_MapToUnitState:
_stUnit.bComm		:= _bComm AND NOT _stReadMap.nPcsStatus.5;
_stUnit.bFault		:= _stReadMap.nPcsStatus.1;
_stUnit.bCtrlReady	:= _stReadMap.nRemoteMode = 1;

IF NOT _stUnit.bComm THEN
	_stUnit.eRunState := E_RunState.Unknown;
ELSIF _stUnit.bFault THEN
	_stUnit.eRunState := E_RunState.Fault;
ELSIF NOT _stReadMap.nPcsStatus.0 THEN
	_stUnit.eRunState := E_RunState.Stop;
ELSIF _bStandbyMode THEN
	_stUnit.eRunState := E_RunState.Standby;
ELSE
	_stUnit.eRunState := E_RunState.Run;
END_IF

_stUnit.stP.fValue	:= INT_TO_REAL(_stReadMap.nAcActive) * 0.1 * SEL(i_bPInvert, 1.0, -1.0);
_stUnit.stP.bValid	:= _stUnit.bComm;
_stUnit.stQ.fValue	:= INT_TO_REAL(_stReadMap.nAcReactive) * 0.1;
_stUnit.stQ.bValid	:= _stUnit.bComm;
END_ACTION

ACTION A_ReadRegisters:
// 읽기 주기마다 한 번 (Helios A_ReadPcsData와 같은 순서)
IF NOT _bReading THEN
	IF _bReadDue THEN
		_fbMbRead(sIPAddr := i_sIpAddr, nTCPPort := i_nPort, nUnitID := i_nUnitId,
				nQuantity := SIZEOF(_stReadMap) / 2, nMBAddr := 1, cbLength := SIZEOF(_stReadMap),
				pDestAddr := ADR(_stReadMap), tTimeout := i_tTimeout, bExecute := TRUE);
		_bReading := TRUE;
	END_IF
ELSE
	_fbMbRead(bExecute := FALSE);
	IF NOT _fbMbRead.bBusy THEN
		_bReadError	:= _fbMbRead.bError;
		_nReadErrId	:= _fbMbRead.nErrId;
		IF NOT _fbMbRead.bError THEN
			M_MarkAlive();
		END_IF
		_bReading := FALSE;
	END_IF
END_IF
END_ACTION

ACTION A_WriteQueue:
CASE _nWriteStep OF
	0:	// 다음 일: 상태 명령이 먼저, 그다음 출력
		_nSendCount := 0;
		IF _nCmdRegCount > 0 THEN
			FOR _nCopyIdx := 1 TO _nCmdRegCount DO
				_anSendAddr[_nCopyIdx]	:= _anCmdRegAddr[_nCopyIdx];
				_anSendValue[_nCopyIdx]	:= _anCmdRegValue[_nCopyIdx];
			END_FOR
			_nSendCount := _nCmdRegCount;
			_nCmdRegCount := 0;
		ELSIF _bPowerPending THEN
			IF _nPowerDir <> 0 AND _nPowerDir <> _nDirWritten THEN
				_anSendAddr[1] := 106;	_anSendValue[1] := 1;
				_anSendAddr[2] := 103;	_anSendValue[2] := _nPowerDir;
				_anSendAddr[3] := 107;	_anSendValue[3] := _nPowerAbs;
				_nSendCount := 3;
			ELSE
				_anSendAddr[1] := 107;	_anSendValue[1] := _nPowerAbs;
				_nSendCount := 1;
			END_IF
			_bPowerPending := FALSE;
		END_IF
		IF _nSendCount > 0 THEN
			_nSendIdx	:= 1;
			_nWriteStep	:= 1;
		END_IF

	1:	// 레지스터 하나 쓰기 시작
		_fbMbWrite(sIPAddr := i_sIpAddr, nTCPPort := i_nPort, nUnitID := i_nUnitId,
				 nQuantity := 1, nMBAddr := _anSendAddr[_nSendIdx], cbLength := 2,
				 pSrcAddr := ADR(_anSendValue[_nSendIdx]), tTimeout := i_tTimeout, bExecute := TRUE);
		_nWriteStep := 2;

	2:	// 끝나기 기다림
		_fbMbWrite(bExecute := FALSE);
		IF NOT _fbMbWrite.bBusy THEN
			_bWriteError := _fbMbWrite.bError;
			_nWriteErrId := _fbMbWrite.nErrId;
			IF NOT _fbMbWrite.bError AND _anSendAddr[_nSendIdx] = 103 THEN
				_nDirWritten := _anSendValue[_nSendIdx];
			END_IF
			IF _fbMbWrite.bError THEN
				_nSendIdx := _nSendCount;		// 실패하면 이 일은 그만 (상태 명령은 시퀀서가 다시 보냄)
			END_IF
			_nWriteStep := 3;
		END_IF

	3:	// 간격
		_tonWriteGap(IN := TRUE, PT := i_tWriteGap);
		IF _tonWriteGap.Q THEN
			_tonWriteGap(IN := FALSE);
			IF _nSendIdx < _nSendCount THEN
				_nSendIdx	:= _nSendIdx + 1;
				_nWriteStep	:= 1;
			ELSE
				_nWriteStep	:= 0;
			END_IF
		END_IF
END_CASE
END_ACTION

METHOD M_Cycle
_bReadDue := M_IsReadTime();
A_ReadRegisters();
M_UpdateComm();
A_MapToUnitState();
A_WriteQueue();
END_METHOD

METHOD M_GetUnitState : ST_UnitState
VAR_INPUT
	i_nSub		: UINT;
END_VAR
IF i_nSub = 1 THEN
	M_GetUnitState := _stUnit;
END_IF
END_METHOD

METHOD PRIVATE M_QueueCmdAndApply		// 상태 명령 보낼 목록을 새로 만듦: 명령 레지스터 하나 + 적용 신호(105 ← 1)
VAR_INPUT
	i_nAddr		: UINT;
	i_nValue	: INT;
END_VAR
_nCmdRegCount := 0;
M_QueueRegister(i_nAddr, i_nValue);
M_QueueRegister(105, 1);
END_METHOD

METHOD PRIVATE M_QueueRegister		// 상태 명령 보낼 목록에 레지스터 하나(주소 ← 값) 추가
VAR_INPUT
	i_nAddr		: UINT;
	i_nValue	: INT;
END_VAR
IF _nCmdRegCount < 5 THEN
	_nCmdRegCount := _nCmdRegCount + 1;
	_anCmdRegAddr[_nCmdRegCount]	:= i_nAddr;
	_anCmdRegValue[_nCmdRegCount]	:= i_nValue;
END_IF
END_METHOD

METHOD M_SetPower : BOOL
VAR_INPUT
	i_nSub		: UINT;
	i_fP		: REAL;			// kW, 방전 +
	i_fQ		: REAL;			// 이 맵에는 Q 지령이 없음
END_VAR
IF i_nSub <> 1 THEN
	RETURN;
END_IF
IF i_fP > 0.05 THEN
	_nPowerDir := 2;			// 방전
ELSIF i_fP < -0.05 THEN
	_nPowerDir := 1;			// 충전
ELSE
	_nPowerDir := 0;			// 0 kW: 방향은 그대로 두고 107만
END_IF
// [결함 13 수정 2026-11-04: 지령·배율이 숫자가 아니면 0 (LIMIT·REAL_TO_INT에서 FPU 예외). 원래 _nPowerAbs := REAL_TO_INT(LIMIT(0.0, ABS(i_fP) * i_fPScale, 32767.0));]
IF F_RealOk(i_fP) AND F_RealOk(i_fPScale) THEN
	_nPowerAbs	:= REAL_TO_INT(LIMIT(0.0, ABS(i_fP) * i_fPScale, 32767.0));
ELSE
	_nPowerAbs	:= 0;
END_IF
_bPowerPending	:= TRUE;
M_SetPower := TRUE;
END_METHOD

METHOD M_SetStateCmd : BOOL
VAR_INPUT
	i_nSub		: UINT;
	i_stCmd		: ST_PcsCmd;
END_VAR
IF i_nSub <> 1 THEN
	RETURN;
END_IF

CASE i_stCmd.eCmd OF
	E_PcsCmd.Run:
		_bStandbyMode := FALSE;
		_nDirWritten := 0;			// 첫 출력 때 방향(103)을 다시 씀
		IF _stUnit.eRunState = E_RunState.Stop THEN
			M_QueueCmdAndApply(101, 55);			// 기동
		END_IF
		// 이미 운전 중이면 쓸 것 없음: Run으로 보고하고 출력 지령을 따름

	E_PcsCmd.Standby:
		_bStandbyMode := TRUE;
		_nCmdRegCount := 0;
		IF _stUnit.eRunState = E_RunState.Stop THEN
			M_QueueRegister(101, 55);
			M_QueueRegister(105, 1);
		END_IF
		M_QueueRegister(106, 1);
		M_QueueRegister(103, 0);
		M_QueueRegister(107, 0);

	E_PcsCmd.Stop,
	E_PcsCmd.EStop:
		_bStandbyMode := FALSE;
		_nDirWritten := 0;
		M_QueueCmdAndApply(101, 99);

	E_PcsCmd.Reset:
		M_QueueCmdAndApply(102, 33);
ELSE
	RETURN;
END_CASE
M_SetStateCmd := TRUE;
END_METHOD

PROPERTY RawMap : ST_PlaspoPcsRaw		// 마지막으로 읽은 레지스터 맵 (보고 매핑용. 제어에 쓰지 않음)
GET
RawMap := _stReadMap;
END_GET
END_PROPERTY

END_FUNCTION_BLOCK

// ---- 20_Module/Virtual/FB_PcsSim.TcPOU
FUNCTION_BLOCK FB_PcsSim EXTENDS FB_DeviceBase IMPLEMENTS I_Pcs		// 가상 PCS (시험용)
VAR_INPUT
	i_tTau			: TIME := T#500MS;	// 출력 응답 시정수
	i_bForceFault	: BOOL;				// 시험: 전 유닛 고장
	i_bForceLocal	: BOOL;				// 시험: 로컬 모드 (PMS 제어 불가)
	i_bForceCommLoss	: BOOL;			// 시험: 통신 끊김 (응답 안 함. i_tCommTimeout 뒤 통신 이상)
	i_bIgnoreCmd	: BOOL;				// 시험: 상태 명령을 접수하되 상태는 바꾸지 않음 (P/Q 지령은 적용)
	i_bFaultFlagOnly	: BOOL;			// 시험: 운전 상태는 그대로 두고 고장 표시만 켬 (해제도 이 입력으로 함)
END_VAR
VAR
	_aeState		: ARRAY[1..GVL_PARAM.MAX_SUB] OF E_RunState;
	_afPSet			: ARRAY[1..GVL_PARAM.MAX_SUB] OF REAL;
	_afQSet			: ARRAY[1..GVL_PARAM.MAX_SUB] OF REAL;
	_afbPLag			: ARRAY[1..GVL_PARAM.MAX_SUB] OF FB_Lpf;
	_afbQLag			: ARRAY[1..GVL_PARAM.MAX_SUB] OF FB_Lpf;
	_astUnit		: ARRAY[1..GVL_PARAM.MAX_SUB] OF ST_UnitState;
END_VAR

METHOD M_Cycle
VAR
	u		: UINT;
	fPTarget		: REAL;
	fQTarget		: REAL;
END_VAR
IF M_IsReadTime() AND NOT i_bForceCommLoss THEN		// 읽기 주기마다 응답한 것으로 봄 (시험: 통신 끊김이면 응답 안 함)
	M_MarkAlive();
END_IF
M_UpdateComm();

FOR u := 1 TO GVL_PARAM.MAX_SUB DO
	IF _aeState[u] = E_RunState.Unknown THEN
		_aeState[u] := E_RunState.Stop;
	END_IF
	IF i_bForceFault THEN
		_aeState[u] := E_RunState.Fault;
	END_IF

	// 운전 중이면 지령을, 아니면 0을 1차 지연으로 따라감
	IF _aeState[u] = E_RunState.Run THEN
		fPTarget := _afPSet[u];
		fQTarget := _afQSet[u];
	ELSE
		fPTarget := 0;
		fQTarget := 0;
	END_IF
	_afbPLag[u](i_fIn := fPTarget, i_tTau := i_tTau);
	_afbQLag[u](i_fIn := fQTarget, i_tTau := i_tTau);

	_astUnit[u].bComm		:= _bComm;
	_astUnit[u].eRunState	:= _aeState[u];
	_astUnit[u].bCtrlReady	:= NOT i_bForceLocal;
	_astUnit[u].bFault		:= (_aeState[u] = E_RunState.Fault) OR i_bFaultFlagOnly;
	_astUnit[u].stP.fValue	:= _afbPLag[u].q_fOut;
	_astUnit[u].stP.bValid	:= TRUE;
	_astUnit[u].stQ.fValue	:= _afbQLag[u].q_fOut;
	_astUnit[u].stQ.bValid	:= TRUE;
END_FOR
END_METHOD

METHOD M_GetUnitState : ST_UnitState
VAR_INPUT
	i_nSub		: UINT;
END_VAR
IF i_nSub >= 1 AND i_nSub <= GVL_PARAM.MAX_SUB THEN
	M_GetUnitState := _astUnit[i_nSub];
END_IF
END_METHOD

METHOD M_SetPower : BOOL
VAR_INPUT
	i_nSub		: UINT;
	i_fP		: REAL;
	i_fQ		: REAL;
END_VAR
IF i_nSub < 1 OR i_nSub > GVL_PARAM.MAX_SUB THEN
	RETURN;
END_IF
_afPSet[i_nSub] := i_fP;
_afQSet[i_nSub] := i_fQ;
M_SetPower := TRUE;
END_METHOD

METHOD M_SetStateCmd : BOOL
VAR_INPUT
	i_nSub		: UINT;
	i_stCmd		: ST_PcsCmd;
END_VAR
IF i_nSub < 1 OR i_nSub > GVL_PARAM.MAX_SUB THEN
	RETURN;
END_IF

CASE i_stCmd.eCmd OF
	E_PcsCmd.Run:
		IF NOT i_bIgnoreCmd AND _aeState[i_nSub] <> E_RunState.Fault THEN _aeState[i_nSub] := E_RunState.Run; END_IF

	E_PcsCmd.Standby:
		IF NOT i_bIgnoreCmd AND _aeState[i_nSub] <> E_RunState.Fault THEN _aeState[i_nSub] := E_RunState.Standby; END_IF

	E_PcsCmd.Stop,
	E_PcsCmd.EStop:
		IF NOT i_bIgnoreCmd AND _aeState[i_nSub] <> E_RunState.Fault THEN _aeState[i_nSub] := E_RunState.Stop; END_IF

	E_PcsCmd.Reset:
		IF NOT i_bIgnoreCmd AND _aeState[i_nSub] = E_RunState.Fault AND NOT i_bForceFault THEN _aeState[i_nSub] := E_RunState.Stop; END_IF
ELSE
	RETURN;		// 배터리 명령 등은 PCS가 받지 않음
END_CASE

M_SetStateCmd := TRUE;
END_METHOD

END_FUNCTION_BLOCK

// ---- 20_Module/Report/FB_RptPlaspoPcs.TcPOU
FUNCTION_BLOCK FB_RptPlaspoPcs		// 보고 매핑: 플라스포 PCS 읽기값 + 코어 결과 → MQTT pcs 발행 레코드 (보고 전용, 제어에 쓰지 않음)
(* 필드 대응 (플라스포 읽기 맵 ST_PlaspoPcsRaw, 괄호는 레지스터 번호):
   SystemOperationMode  코어 운전 모드 (Manual 0, Auto 1)
   OperationMode        nOpMode (4) 그대로
   PMSActivePower       PMS가 이 PCS에 낸 지령 kW (분배 결과. 장비 쓰기를 막아도 나옴)
   RemoteMode           nRemoteMode (3)
   Status               nPcsStatus (1) 그대로: bit0 운전, bit1 고장, bit2 경고, bit5 PCS 내부 통신 이상
   AcActivePower·AcReactivePower  드라이버가 변환한 P·Q (방전 +, 0.1 kW·kvar)
   PowerFactor          nAcPf (29) × i_fPfScale
   Frequency            nAcFreq (26) × 0.1
   AcRs·St·TrVoltage    anAcVolt[1..3] (20~22) × i_fVoltScale  (선간 전압으로 가정)
   AcR·S·TVoltage       읽지 않음 → 0
   AcR·S·TCurrent       anAcCurrent[1..3] (23~25) × i_fCurrScale
   DcLinkVoltage·DcVoltage  nDcLinkVolt (36)·nDcVolt (37) × i_fDcVoltScale
   DcCurrent            nDcCurrent (38) × i_fDcCurrScale
   DcActivePower        nDcPower (39) × i_fDcPowerScale
   InsulationResistance 읽지 않음 → 0
   Temperature1~4       anIgbtTemp[1..4] (12~15) × i_fTempScale
   Temperature5~8       anAcFilterTemp[1..4] (16~19) × i_fTempScale
   Warning1             anFault[5] (11). Warning2~10 → 0
   Fault1~4             anFault[1..4] (7~10). Fault5~10 → 0
   통신이 끊기면 레코드 전체가 0 (이 값만으로는 끊김을 알 수 없으니 GVL_IF.g_stReport.abPcsComm을 봄)
   배율(i_f…Scale)은 레지스터 맵 문서로 확인되지 않은 값이라 기본 1.0 (= 레지스터 값 그대로). 실제 값과 비교해 맞출 것 *)
VAR_INPUT
	i_stRaw			: ST_PlaspoPcsRaw;	// 드라이버 FB_PlaspoPcs.RawMap
	i_stUnit		: ST_UnitState;		// 이 PCS의 유닛 상태 (FB_Snapshot)
	i_eOpMode		: E_OpMode;			// 이 유닛의 실제 운전 모드 (FB_ModeSwitch)
	i_fPCmd			: REAL;				// kW, PMS가 낸 지령 (FB_Distributor 유닛 지령)
	i_fPfScale		: REAL := 1.0;
	i_fVoltScale	: REAL := 1.0;
	i_fCurrScale	: REAL := 1.0;
	i_fDcVoltScale	: REAL := 1.0;
	i_fDcCurrScale	: REAL := 1.0;
	i_fDcPowerScale	: REAL := 1.0;
	i_fTempScale	: REAL := 1.0;
END_VAR
VAR_OUTPUT
	q_stPcs			: ST_PcsPublish_V1;	// 발행 직전 레코드 (DeviceIndex는 PRG_Mqtt가 채움)
	q_bComm			: BOOL;				// 통신 정상
END_VAR
VAR
	_stNone			: ST_PcsPublish_V1;
END_VAR

q_stPcs := _stNone;
q_bComm := i_stUnit.bComm;
IF NOT q_bComm THEN
	RETURN;
END_IF

IF i_eOpMode = E_OpMode.Auto THEN
	q_stPcs.SystemOperationMode := 1;
ELSE
	q_stPcs.SystemOperationMode := 0;
END_IF
q_stPcs.OperationMode		:= UINT_TO_UDINT(i_stRaw.nOpMode);
q_stPcs.PMSActivePower		:= i_fPCmd;
q_stPcs.RemoteMode			:= UINT_TO_UDINT(i_stRaw.nRemoteMode);
q_stPcs.Status				:= DWORD_TO_UDINT(WORD_TO_DWORD(i_stRaw.nPcsStatus));

q_stPcs.AcActivePower		:= i_stUnit.stP.fValue;
q_stPcs.AcReactivePower		:= i_stUnit.stQ.fValue;
q_stPcs.PowerFactor			:= INT_TO_REAL(i_stRaw.nAcPf) * i_fPfScale;
q_stPcs.Frequency			:= UINT_TO_REAL(i_stRaw.nAcFreq) * 0.1;

q_stPcs.AcRsVoltage			:= UINT_TO_REAL(i_stRaw.anAcVolt[1]) * i_fVoltScale;
q_stPcs.AcStVoltage			:= UINT_TO_REAL(i_stRaw.anAcVolt[2]) * i_fVoltScale;
q_stPcs.AcTrVoltage			:= UINT_TO_REAL(i_stRaw.anAcVolt[3]) * i_fVoltScale;
q_stPcs.AcRCurrent			:= UINT_TO_REAL(i_stRaw.anAcCurrent[1]) * i_fCurrScale;
q_stPcs.AcSCurrent			:= UINT_TO_REAL(i_stRaw.anAcCurrent[2]) * i_fCurrScale;
q_stPcs.AcTCurrent			:= UINT_TO_REAL(i_stRaw.anAcCurrent[3]) * i_fCurrScale;

q_stPcs.DcLinkVoltage		:= UINT_TO_REAL(i_stRaw.nDcLinkVolt) * i_fDcVoltScale;
q_stPcs.DcVoltage			:= UINT_TO_REAL(i_stRaw.nDcVolt) * i_fDcVoltScale;
q_stPcs.DcCurrent			:= INT_TO_REAL(i_stRaw.nDcCurrent) * i_fDcCurrScale;
q_stPcs.DcActivePower		:= INT_TO_REAL(i_stRaw.nDcPower) * i_fDcPowerScale;

q_stPcs.Temperature1		:= INT_TO_REAL(i_stRaw.anIgbtTemp[1]) * i_fTempScale;
q_stPcs.Temperature2		:= INT_TO_REAL(i_stRaw.anIgbtTemp[2]) * i_fTempScale;
q_stPcs.Temperature3		:= INT_TO_REAL(i_stRaw.anIgbtTemp[3]) * i_fTempScale;
q_stPcs.Temperature4		:= INT_TO_REAL(i_stRaw.anIgbtTemp[4]) * i_fTempScale;
q_stPcs.Temperature5		:= INT_TO_REAL(i_stRaw.anAcFilterTemp[1]) * i_fTempScale;
q_stPcs.Temperature6		:= INT_TO_REAL(i_stRaw.anAcFilterTemp[2]) * i_fTempScale;
q_stPcs.Temperature7		:= INT_TO_REAL(i_stRaw.anAcFilterTemp[3]) * i_fTempScale;
q_stPcs.Temperature8		:= INT_TO_REAL(i_stRaw.anAcFilterTemp[4]) * i_fTempScale;

q_stPcs.Warning1			:= DWORD_TO_UDINT(WORD_TO_DWORD(i_stRaw.anFault[5]));
q_stPcs.Fault1				:= DWORD_TO_UDINT(WORD_TO_DWORD(i_stRaw.anFault[1]));
q_stPcs.Fault2				:= DWORD_TO_UDINT(WORD_TO_DWORD(i_stRaw.anFault[2]));
q_stPcs.Fault3				:= DWORD_TO_UDINT(WORD_TO_DWORD(i_stRaw.anFault[3]));
q_stPcs.Fault4				:= DWORD_TO_UDINT(WORD_TO_DWORD(i_stRaw.anFault[4]));

END_FUNCTION_BLOCK

// ---- 20_Module/Driver/Esolution/FB_EsolutionBms.TcPOU
FUNCTION_BLOCK FB_EsolutionBms EXTENDS FB_DeviceBase IMPLEMENTS I_Bms

VAR_INPUT
	i_bEnable : BOOL;
	i_sIpAddr : STRING(15);
	i_nPort : UINT := 502;
	i_nUnitId : BYTE := 1;
	i_tTimeout : TIME := T#1S;
	i_bWritePermit : BOOL; // site dispatcher: config OK AND active PLC
END_VAR
VAR_OUTPUT
	q_eRequestResult : E_UpsResult;
	q_nTransportError : UDINT;
END_VAR
VAR
	_fbJob : FB_UpsModbusJob;
	_bLaunch : BOOL;
	_bCurrentWrite : BOOL;
	_bDiscardResponse : BOOL; // response started before a disable must not complete a new snapshot
	_nFunction : UINT;
	_nAddress : WORD;
	_nQuantity : WORD;
	_wValue : WORD;
	_bPendingWrite : BOOL;
	_nPendingAddress : WORD;
	_wPendingValue : WORD;
	_nPendingQty : WORD; // 1 = FC06, 2~3 = FC16 같은 값 여러 칸 [2026-11-13]
	_awValues : ARRAY[0..2] OF WORD;
	_nPoll : UINT;
	_nCopy : UINT;
	_bReadDue : BOOL;
	_bCycle : BOOL; // 2026-11-23 기본 한 바퀴(시스템·랙 아날로그·랙 상태 3개) 읽는 중 (명세 DV-04 v2.46)
	_bDetailReq : BOOL; // 랙 상세 한 조각을 읽을 차례
	_tonDetailRead : TON; // 랙 상세 읽기 간격
END_VAR

VAR_INPUT
	i_nRackCount : UINT := 1; // configure actual installed count, max10
	i_nModuleCount : UINT := GVL_PARAM.MODULES_PER_RACK; // installed modules; map stride remains 17 slots
	i_bReadDetails : BOOL := FALSE; // enable after unused module-slot response is confirmed
	i_tHeartbeatTimeout : TIME := T#10S;
	i_tDetailTimeout : TIME := T#60S;
	i_tDetailPeriod : TIME := T#100MS; // 랙 상세 한 조각(125 레지스터) 읽는 간격. 기본 한 바퀴(i_tReadPeriod) 사이사이에 읽음 (명세 DV-04 v2.46)
	i_stTime : ST_LocalTime; // PMS 현지 시각 (MAIN.fbClock). BMS 시각 동기용 (명세 WR-BAT-01 v2.35)
	i_tTimeSync : TIME := T#1H; // BMS 시각 동기 주기 (BAT 질의 Q1: 1시간). T#0S = 끔
END_VAR
VAR_OUTPUT
	q_stRaw : ST_EsolutionRaw;
	q_stState : ST_EsolutionState;
	q_nTimeSyncCount : UDINT; // 시각 동기 쓰기를 넣은 횟수 (HR 40005~40007)
END_VAR
VAR
	_stWork : ST_EsolutionRaw;
	_stBat : ST_BatState;
	_nSampleSeq : UDINT;
	_nRack : UINT;
	_nOffset : UINT;
	_nDetailRack : UINT := 1;
	_nDetailOffset : UINT;
	_nDetailChunk : UINT;
	_wHeartbeat : WORD;
	_bHeartbeatChanged : BOOL;
	_tonHeartbeat : TON;
	_atonDetail : ARRAY[1..10] OF TON;
	_abDetailUpdated : ARRAY[1..10] OF BOOL;
	_wInstalledMask : WORD;
	_nLastRackCount : UINT;
	_nLastCoreCmdSeq : UDINT;
	_bHaveCoreCmd : BOOL;
	_tonTimeSync : TON;
	_bTimeSyncDue : BOOL := TRUE; // 통신이 붙으면 먼저 한 번
	_awPendingValues : ARRAY[0..2] OF WORD; // FC16 칸별 값 (보통은 셋 다 같은 값, 시각 동기만 다름)
END_VAR

PROPERTY BatState : ST_BatState
GET
BatState:=_stBat;
END_GET
END_PROPERTY

METHOD M_CheckSet : WSTRING(63)
M_CheckSet:="";
IF i_bEnable THEN
	IF i_sIpAddr='' OR i_nPort=0 THEN M_CheckSet:="TCP endpoint missing";
	ELSIF i_tReadPeriod<=T#0MS OR i_tTimeout<=T#0MS OR i_tCommTimeout<=i_tReadPeriod THEN M_CheckSet:="Invalid timing";
	END_IF
END_IF
IF i_nRackCount<1 OR i_nRackCount>10 OR i_nModuleCount<1 OR i_nModuleCount>17 THEN
	M_CheckSet:="Rack/module range";
END_IF
END_METHOD

METHOD M_Cycle
_bReadDue := M_IsReadTime();
IF _bReadDue THEN _bCycle:=TRUE; END_IF // 기본 한 바퀴 시작 (명세 DV-04 v2.46: 주기 = 한 바퀴)
_tonDetailRead(IN:=i_bReadDetails AND NOT _tonDetailRead.Q, PT:=i_tDetailPeriod);
IF _tonDetailRead.Q THEN _bDetailReq:=TRUE; END_IF
IF NOT i_bEnable THEN
	_bDiscardResponse:=_bDiscardResponse OR _fbJob.q_bBusy;
	_bLaunch:=FALSE;
END_IF
IF NOT i_bEnable OR NOT i_bWritePermit OR NOT GVL_PARAM.UPS_CONTROL_ENABLED THEN
	_bPendingWrite := FALSE;
	// A queued but not yet started FC06 must not survive a gate transition.
	IF _bLaunch AND _bCurrentWrite THEN _bLaunch := FALSE; END_IF
END_IF
_fbJob(i_sIpAddr:=i_sIpAddr,i_nPort:=i_nPort,i_nUnitId:=i_nUnitId,i_tTimeout:=i_tTimeout,
	i_bExecute:=_bLaunch,i_bWritePermit:=i_bWritePermit AND i_bEnable,
	i_nFunction:=_nFunction,i_nAddress:=_nAddress,i_nQuantity:=_nQuantity,i_wValue:=_wValue,i_awValues:=_awValues);
_bLaunch := FALSE;
IF _fbJob.q_bDone THEN
	q_nTransportError := _fbJob.q_nErrorId;
	IF _bCurrentWrite THEN M_MarkWriteResult(NOT _fbJob.q_bError); END_IF
END_IF

IF i_nRackCount<1 OR i_nRackCount>10 OR i_nModuleCount<1 OR i_nModuleCount>17 THEN
	_bLaunch:=FALSE; _bPendingWrite:=FALSE;
	q_stState.bComm:=FALSE; q_stState.bValid:=FALSE; _stBat.bComm:=FALSE;
	RETURN;
END_IF
IF _nLastRackCount<>i_nRackCount THEN
	_nLastRackCount:=i_nRackCount; _nDetailRack:=1; _nDetailOffset:=0;
	FOR _nRack:=1 TO 10 DO q_stState.abDetailValid[_nRack]:=FALSE; END_FOR
END_IF
_bHeartbeatChanged:=FALSE;
FOR _nRack:=1 TO 10 DO _abDetailUpdated[_nRack]:=FALSE; END_FOR
IF _fbJob.q_bDone AND _bDiscardResponse THEN
	_bDiscardResponse:=FALSE; _nPoll:=0; _bCycle:=FALSE; _bDetailReq:=FALSE;
ELSIF _fbJob.q_bDone AND NOT _bCurrentWrite THEN
	IF _fbJob.q_bError THEN
		IF _nPoll=3 THEN _nDetailOffset:=0; _bDetailReq:=FALSE; ELSE _bCycle:=FALSE; END_IF // 다음 차례에 다시
		_nPoll:=0;
	ELSE
		CASE _nPoll OF
			0: FOR _nCopy:=0 TO 26 DO _stWork.awSystem[_nCopy]:=_fbJob.q_awData[_nCopy]; END_FOR
			1: FOR _nCopy:=0 TO 39 DO _stWork.awRackAnalog[_nCopy]:=_fbJob.q_awData[_nCopy]; END_FOR
			2:
				FOR _nCopy:=0 TO 89 DO _stWork.awRackStatus[_nCopy]:=_fbJob.q_awData[_nCopy]; END_FOR
				q_stRaw.awSystem:=_stWork.awSystem;
				q_stRaw.awRackAnalog:=_stWork.awRackAnalog;
				q_stRaw.awRackStatus:=_stWork.awRackStatus;
				_bHeartbeatChanged:=_nSampleSeq=0 OR _wHeartbeat<>q_stRaw.awSystem[0];
				_wHeartbeat:=q_stRaw.awSystem[0]; _nSampleSeq:=F_UpsNextSeq(_nSampleSeq); M_MarkAlive();
			3:
				FOR _nCopy:=0 TO _nDetailChunk-1 DO
					_stWork.aawDetail[_nDetailRack,_nDetailOffset+_nCopy]:=_fbJob.q_awData[_nCopy];
				END_FOR
				IF _nDetailOffset+_nDetailChunk=406 THEN
					FOR _nCopy:=0 TO 405 DO q_stRaw.aawDetail[_nDetailRack,_nCopy]:=_stWork.aawDetail[_nDetailRack,_nCopy]; END_FOR
					q_stState.anDetailSeq[_nDetailRack]:=F_UpsNextSeq(q_stState.anDetailSeq[_nDetailRack]);
					_abDetailUpdated[_nDetailRack]:=TRUE;
					q_stState.abDetailValid[_nDetailRack]:=TRUE;
					_nDetailOffset:=0;
					IF _nDetailRack>=i_nRackCount THEN _nDetailRack:=1; ELSE _nDetailRack:=_nDetailRack+1; END_IF
				ELSE _nDetailOffset:=_nDetailOffset+_nDetailChunk; END_IF
		END_CASE
		IF _nPoll=2 THEN _nPoll:=0; _bCycle:=FALSE; // 기본 한 바퀴 끝
		ELSIF _nPoll=3 THEN _nPoll:=0; _bDetailReq:=FALSE; // 랙 상세 한 조각 끝
		ELSE _nPoll:=_nPoll+1; END_IF
	END_IF
END_IF
M_UpdateComm();
_tonHeartbeat(IN:=NOT _bHeartbeatChanged,PT:=i_tHeartbeatTimeout);
// System Data 1~27
q_stState.nHeartbeat:=q_stRaw.awSystem[0]; // 1. 하트비트
q_stState.fVoltageV:=WORD_TO_REAL(q_stRaw.awSystem[1])*0.1; // 2. 전체 전압 (V)
q_stState.fCurrentA:=F_UpsSignedWord(q_stRaw.awSystem[2])*0.1; // 3. 전체 전류 (A)
q_stState.fSocPct:=WORD_TO_REAL(q_stRaw.awSystem[3])*0.1; // 4. 충전 상태 (%)
q_stState.fSohPct:=WORD_TO_REAL(q_stRaw.awSystem[4]); // 5. 건강 상태 (%)
q_stState.fChargePowerKw:=WORD_TO_REAL(q_stRaw.awSystem[5]); // 6. 충전 전력 (kW)
q_stState.fDischargePowerKw:=WORD_TO_REAL(q_stRaw.awSystem[6]); // 7. 방전 전력 (kW)
q_stState.fMaxCellVoltageMv:=WORD_TO_REAL(q_stRaw.awSystem[7]); // 8. 최대 셀 전압 (mV)
q_stState.fMinCellVoltageMv:=WORD_TO_REAL(q_stRaw.awSystem[8]); // 9. 최소 셀 전압 (mV)
q_stState.fAvgCellVoltageMv:=WORD_TO_REAL(q_stRaw.awSystem[9]); // 10. 평균 셀 전압 (mV)
q_stState.nMaxCellVoltageLocation:=q_stRaw.awSystem[10]; // 11. 최대 셀 전압 위치
q_stState.nMinCellVoltageLocation:=q_stRaw.awSystem[11]; // 12. 최소 셀 전압 위치
q_stState.fMaxCellTemperatureC:=F_UpsSignedWord(q_stRaw.awSystem[12])*0.1; // 13. 최고 셀 온도 (℃)
q_stState.fMinCellTemperatureC:=F_UpsSignedWord(q_stRaw.awSystem[13])*0.1; // 14. 최저 셀 온도 (℃)
q_stState.fAvgCellTemperatureC:=F_UpsSignedWord(q_stRaw.awSystem[14])*0.1; // 15. 평균 셀 온도 (℃)
q_stState.nMaxCellTemperatureLocation:=q_stRaw.awSystem[15]; // 16. 최고 셀 온도 위치
q_stState.nMinCellTemperatureLocation:=q_stRaw.awSystem[16]; // 17. 최저 셀 온도 위치
q_stState.fMaxRackSocPct:=WORD_TO_REAL(q_stRaw.awSystem[17])*0.1; // 18. 최대 랙 SOC (%)
q_stState.fMinRackSocPct:=WORD_TO_REAL(q_stRaw.awSystem[18])*0.1; // 19. 최소 랙 SOC (%)
q_stState.fMaxRackVoltageV:=WORD_TO_REAL(q_stRaw.awSystem[19])*0.1; // 20. 최대 랙 전압 (V)
q_stState.fMinRackVoltageV:=WORD_TO_REAL(q_stRaw.awSystem[20])*0.1; // 21. 최소 랙 전압 (V)
q_stState.fChargeLimitKw:=WORD_TO_REAL(q_stRaw.awSystem[21]); // 22. 충전 허용 전력 (kW)
q_stState.fDischargeLimitKw:=WORD_TO_REAL(q_stRaw.awSystem[22]); // 23. 방전 허용 전력 (kW)
q_stState.fChargeCurrentLimitA:=WORD_TO_REAL(q_stRaw.awSystem[23]); // 24. 충전 허용 전류 (A)
q_stState.fDischargeCurrentLimitA:=WORD_TO_REAL(q_stRaw.awSystem[24]); // 25. 방전 허용 전류 (A)
q_stState.wSystemContactor:=q_stRaw.awSystem[25]; // 26. 시스템 컨택터 상태 (맵 v1.4)
q_stState.wRackContactor:=q_stRaw.awSystem[26]; // 27. 랙 컨택터 상태 (맵 v1.4)
q_stState.bChargeContactorClosed:=q_stRaw.awSystem[25].0;
q_stState.bDischargeContactorClosed:=q_stRaw.awSystem[25].1;

q_stState.bComm:=_bComm AND i_bEnable;
q_stState.bFresh:=q_stState.bComm AND NOT _tonHeartbeat.Q;
q_stState.bValid:=q_stState.bFresh AND _nSampleSeq<>0;
q_stState.bWriteFail:=_bWriteFail;
q_stState.nSampleSeq:=_nSampleSeq;
q_stState.nRackCount:=i_nRackCount;
q_stState.nModuleCount:=i_nModuleCount;
q_stState.bWarn:=FALSE; q_stState.bFault:=FALSE; q_stState.bSystemLock:=FALSE;
FOR _nRack:=1 TO 10 DO
	_atonDetail[_nRack](IN:=NOT _abDetailUpdated[_nRack],PT:=i_tDetailTimeout);
	IF _atonDetail[_nRack].Q OR NOT q_stState.bValid OR NOT i_bReadDetails OR _nRack>i_nRackCount THEN
		q_stState.abDetailValid[_nRack]:=FALSE;
	END_IF
	IF _nRack<=i_nRackCount THEN
		_nOffset:=(_nRack-1)*9;
		q_stState.bWarn:=q_stState.bWarn OR (q_stRaw.awRackStatus[_nOffset] AND 16#01FF)<>0
			OR (q_stRaw.awRackStatus[_nOffset+2] AND 16#03FF)<>0 OR q_stRaw.awRackStatus[_nOffset+4].9;
		q_stState.bFault:=q_stState.bFault OR (q_stRaw.awRackStatus[_nOffset+3] AND 16#3FFF)<>0
			OR (q_stRaw.awRackStatus[_nOffset+4] AND 16#05FF)<>0 OR q_stRaw.awRackStatus[_nOffset+5]<>0
			OR (q_stRaw.awRackStatus[_nOffset+6] AND 16#00FF)<>0 OR (q_stRaw.awRackStatus[_nOffset+7] AND 16#8001)<>0;
		q_stState.bSystemLock:=q_stState.bSystemLock OR q_stRaw.awRackStatus[_nOffset].8 OR q_stRaw.awRackStatus[_nOffset+3].13;
	END_IF
END_FOR
// 컨택터 상태는 맵 v1.4 Input 26·27로 판단 (명령이나 운전 모드로 추정하지 않음) [2026-11-13]
// 붙음 = 설치 랙 중 하나라도 붙음 AND 충전·방전 중 하나라도 붙음 (배터리가 버스에 이어짐).
// 그래서 하나라도 붙어 있으면 코어 개방(Open)이 나가고, 개방 확인은 다 떨어져야 됨.
q_stState.bContactorFeedbackKnown:=q_stState.bValid;
_wInstalledMask:=SHL(WORD#1,i_nRackCount)-1;
_stBat.bComm:=q_stState.bValid;
_stBat.bContactorClosed:=q_stState.bValid AND (q_stState.wRackContactor AND _wInstalledMask)<>0
	AND (q_stState.bChargeContactorClosed OR q_stState.bDischargeContactorClosed);
_stBat.bWarn:=q_stState.bWarn; _stBat.bFault:=q_stState.bFault; _stBat.bSysStop:=q_stState.bSystemLock;
_stBat.stSoc.fValue:=q_stState.fSocPct;
_stBat.stSoc.bValid:=q_stState.bValid AND q_stState.fSocPct>=0 AND q_stState.fSocPct<=100;
_stBat.stSoh.fValue:=q_stState.fSohPct;
_stBat.stSoh.bValid:=q_stState.bValid AND q_stState.fSohPct>=0 AND q_stState.fSohPct<=100;
_stBat.fPChgMax:=SEL(q_stState.bValid,0.0,q_stState.fChargeLimitKw);
_stBat.fPDisMax:=SEL(q_stState.bValid,0.0,q_stState.fDischargeLimitKw);
_stBat.bWriteFail:=_bWriteFail;
// BMS 시각 동기 (명세 WR-BAT-01 v2.3·v2.35): HR 40005 YYMM, 40006 DDHH, 40007 mmss (바이트마다 숫자, 예 26년 11월 = 16#1A0B). FC16 한 번
_tonTimeSync(IN:=i_tTimeSync>T#0S AND NOT _tonTimeSync.Q, PT:=i_tTimeSync);
IF _tonTimeSync.Q THEN _bTimeSyncDue:=TRUE; END_IF
IF _bTimeSyncDue AND i_tTimeSync>T#0S AND i_stTime.bValid AND NOT _bPendingWrite THEN
	IF M_QueueWrite(i_nAddress:=4, i_wValue:=SHL(UINT_TO_WORD(i_stTime.nYear MOD 100),8) OR UINT_TO_WORD(i_stTime.nMonth), i_nQuantity:=3) THEN
		_awPendingValues[1]:=SHL(UINT_TO_WORD(i_stTime.nDay),8) OR UINT_TO_WORD(i_stTime.nHour);
		_awPendingValues[2]:=SHL(UINT_TO_WORD(i_stTime.nMinute),8) OR UINT_TO_WORD(i_stTime.nSecond);
		_bTimeSyncDue:=FALSE;
		q_nTimeSyncCount:=q_nTimeSyncCount+1;
	END_IF
END_IF
IF NOT _fbJob.q_bBusy AND NOT _fbJob.q_bDone AND i_bEnable AND i_sIpAddr<>'' THEN
IF _bPendingWrite THEN
	_nAddress:=_nPendingAddress; _nQuantity:=_nPendingQty; _wValue:=_wPendingValue;
	_awValues:=_awPendingValues;
	IF _nPendingQty>1 THEN _nFunction:=16; ELSE _nFunction:=6; END_IF
	_bCurrentWrite:=TRUE; _bPendingWrite:=FALSE; _bLaunch:=TRUE;
ELSIF _bCycle THEN // 기본 한 바퀴: 앞 요청이 끝나면 바로 다음 (명세 DV-04 v2.46)
	_bCurrentWrite:=FALSE;

	_nFunction:=4;
	CASE _nPoll OF
		0: _nAddress:=0; _nQuantity:=27; // 맵 v1.4: 30001~30027
		1: _nAddress:=50; _nQuantity:=40;
		2: _nAddress:=90; _nQuantity:=90;
	END_CASE
	_bLaunch:=TRUE;
ELSIF _bDetailReq AND i_bReadDetails THEN // 랙 상세 한 조각 (기본 한 바퀴 사이사이, i_tDetailPeriod마다)
	_bCurrentWrite:=FALSE;
	_nFunction:=4;
	_nPoll:=3;
	_nDetailChunk:=MIN(125,406-_nDetailOffset);
	_nAddress:=UINT_TO_WORD(500+500*(_nDetailRack-1)+_nDetailOffset);
	_nQuantity:=UINT_TO_WORD(_nDetailChunk);
	_bLaunch:=TRUE;
	END_IF
END_IF
IF NOT i_bEnable THEN _nSampleSeq:=0; _nPoll:=0; _nDetailOffset:=0; _bLaunch:=FALSE; _bCycle:=FALSE; _bDetailReq:=FALSE; END_IF
END_METHOD

METHOD PRIVATE M_QueueWrite : BOOL
VAR_INPUT i_nAddress : WORD; i_wValue : WORD;
	i_nQuantity : WORD; // 1 = FC06. 2~3 = FC16로 i_nAddress부터 같은 값 i_wValue를 여러 칸에 [2026-11-13]
END_VAR
q_eRequestResult := E_UpsResult.Disabled;
IF NOT GVL_PARAM.UPS_CONTROL_ENABLED OR NOT i_bWritePermit OR NOT i_bEnable THEN RETURN; END_IF
	IF i_nQuantity<1 OR i_nQuantity>3 THEN q_eRequestResult := E_UpsResult.BadRequest; RETURN; END_IF
q_eRequestResult := E_UpsResult.CommUnavailable;
	IF NOT q_stState.bValid THEN RETURN; END_IF
q_eRequestResult := E_UpsResult.Busy;
IF _bPendingWrite OR _bCurrentWrite AND (_fbJob.q_bBusy OR _bLaunch) THEN RETURN; END_IF
_nPendingAddress := i_nAddress; _wPendingValue := i_wValue; _nPendingQty := i_nQuantity; _bPendingWrite := TRUE;
_awPendingValues[0] := i_wValue; _awPendingValues[1] := i_wValue; _awPendingValues[2] := i_wValue;	// FC16 같은 값 (시각 동기는 부른 쪽이 1·2칸을 바꿈)
q_eRequestResult := E_UpsResult.Accepted;
M_QueueWrite := TRUE;
END_METHOD

METHOD M_RequestOperation : BOOL
VAR_INPUT i_eOperation : E_EsolutionOperation; END_VAR
IF TO_INT(i_eOperation)<0 OR TO_INT(i_eOperation)>9 THEN q_eRequestResult:=E_UpsResult.Unsupported; RETURN; END_IF
M_RequestOperation:=M_QueueWrite(i_nAddress:=10,i_wValue:=SHL(WORD#1,INT_TO_UINT(TO_INT(i_eOperation))),i_nQuantity:=1);
END_METHOD

METHOD M_SetControl : BOOL
// System protocol v1.4: 0-based holding addresses, uint16 values (NOT 0x55). 하나씩 제어 (EMS command/bat 5~10)
VAR_INPUT i_eControl : E_EsolutionControl; i_bOn : BOOL; END_VAR
CASE i_eControl OF
	E_EsolutionControl.EmergencyShutdown:
		IF NOT i_bOn THEN q_eRequestResult:=E_UpsResult.Unsupported; RETURN; END_IF;
		M_SetControl:=M_QueueWrite(i_nAddress:=11,i_wValue:=1,i_nQuantity:=1);
	E_EsolutionControl.ResetSystem:	// 40031 = 1 (비상차단 해제, 명세 v2.34)
		IF NOT i_bOn THEN q_eRequestResult:=E_UpsResult.Unsupported; RETURN; END_IF;
		M_SetControl:=M_QueueWrite(i_nAddress:=30,i_wValue:=1,i_nQuantity:=1);
	E_EsolutionControl.SystemContactor, E_EsolutionControl.ChargeContactor, E_EsolutionControl.DischargeContactor:
		M_SetControl:=M_QueueWrite(i_nAddress:=INT_TO_WORD(TO_INT(i_eControl)),i_wValue:=BOOL_TO_WORD(i_bOn),i_nQuantity:=1);
ELSE q_eRequestResult:=E_UpsResult.Unsupported;
END_CASE
END_METHOD

METHOD M_SetRackMask : BOOL
// Whole installed-rack bitmap, not an individual-rack pulse. 0 disables ALL installed racks.
VAR_INPUT i_wMask : WORD; END_VAR
IF i_nRackCount<1 OR i_nRackCount>10 THEN q_eRequestResult:=E_UpsResult.BadConfig; RETURN; END_IF
_wInstalledMask:=SHL(WORD#1,i_nRackCount)-1;
IF (i_wMask AND NOT _wInstalledMask)<>0 THEN q_eRequestResult:=E_UpsResult.BadConfig; RETURN; END_IF
M_SetRackMask:=M_QueueWrite(i_nAddress:=0,i_wValue:=i_wMask,i_nQuantity:=1);
END_METHOD

METHOD M_SetStateCmd : BOOL
VAR_INPUT i_stCmd : ST_BatCmd; END_VAR
IF _bHaveCoreCmd AND _nLastCoreCmdSeq=i_stCmd.nSeq THEN
	q_eRequestResult:=E_UpsResult.Duplicate; RETURN;
END_IF
CASE i_stCmd.eCmd OF
	// 투입·개방은 40013(랙 전체)·40014(충전)·40015(방전)를 FC16 한 번에 [1,1,1] / [0,0,0] (2026-11-12 이솔루션 답: 순서 무관, 2026-11-13 사용자 결정 2안)
	E_BatCmd.Close: M_SetStateCmd:=M_QueueWrite(i_nAddress:=INT_TO_WORD(TO_INT(E_EsolutionControl.SystemContactor)),i_wValue:=1,i_nQuantity:=3);
	E_BatCmd.Open: M_SetStateCmd:=M_QueueWrite(i_nAddress:=INT_TO_WORD(TO_INT(E_EsolutionControl.SystemContactor)),i_wValue:=0,i_nQuantity:=3);
	E_BatCmd.EStop: M_SetStateCmd:=M_SetControl(E_EsolutionControl.EmergencyShutdown,TRUE);
	E_BatCmd.Reset: M_SetStateCmd:=M_QueueWrite(i_nAddress:=30,i_wValue:=1,i_nQuantity:=1);
ELSE q_eRequestResult:=E_UpsResult.Unsupported;
END_CASE
IF M_SetStateCmd THEN _bHaveCoreCmd:=TRUE; _nLastCoreCmdSeq:=i_stCmd.nSeq; END_IF
END_METHOD

END_FUNCTION_BLOCK

// ---- 20_Module/Ups/FB_UpsModbusJob.TcPOU
FUNCTION_BLOCK FB_UpsModbusJob
// One latched Modbus transaction. FC03/04 read, FC06 single write, FC16 block write (max 3 words, BMS 40013~40015 [2026-11-13]).
VAR_INPUT
	i_sIpAddr : STRING(15);
	i_nPort : UINT := 502;
	i_nUnitId : BYTE := 1;
	i_tTimeout : TIME := T#1S;
	i_bExecute : BOOL;
	i_bWritePermit : BOOL;
	i_nFunction : UINT;
	i_nAddress : WORD;
	i_nQuantity : WORD;
	i_wValue : WORD;
	i_awValues : ARRAY[0..2] OF WORD; // FC16 values (i_nQuantity words) [2026-11-13]
END_VAR
VAR_OUTPUT
	q_bBusy : BOOL;
	q_bDone : BOOL;
	q_bError : BOOL;
	q_nErrorId : UDINT;
	q_awData : ARRAY[0..124] OF WORD;
END_VAR
VAR
	_fbInput : FB_MBReadInputRegs;
	_fbHolding : FB_MBReadRegs;
	_fbSingle : FB_MBWriteSingleReg;
	_fbMulti : FB_MBWriteRegs; // FC16 [2026-11-13]
	_awValues : ARRAY[0..2] OF WORD;
	_bStartMulti : BOOL;
	_rtExecute : R_TRIG;
	_sIpAddr : STRING(15);
	_nPort : UINT;
	_nUnitId : BYTE;
	_tTimeout : TIME;
	_nAddress : WORD;
	_wValue : WORD;
	_nFunction : UINT;
	_nQuantity : WORD;
	_bStartInput : BOOL;
	_bStartHolding : BOOL;
	_bStartWrite : BOOL;
END_VAR

